ABB RAPID module: Module1.mod

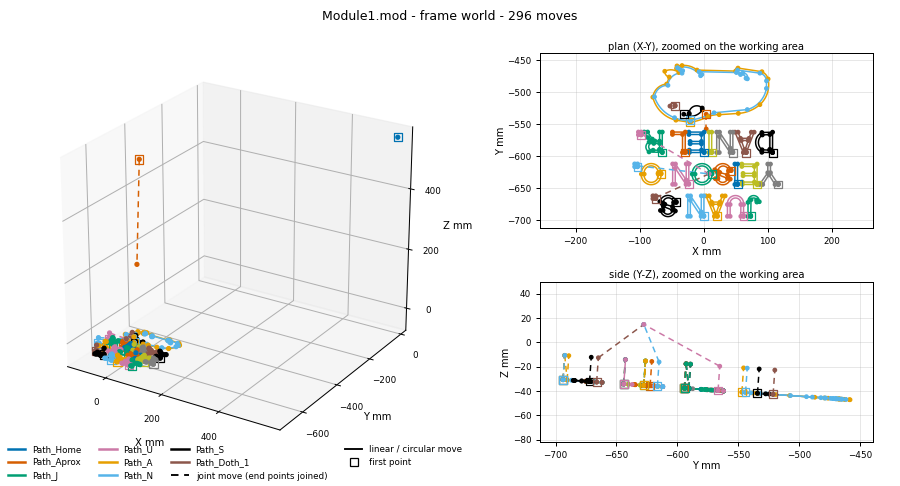
[picture p0: tool path of Module1.mod in frame world, 296 of 313 moves have a stored position in this frame; points joined in program order, loops and branches not executed]
MODULE Module1
    PERS tooldata Tool_Cuy:=[TRUE,[[59.512,0,113],[0.866025404,0,0.5,0]],[1,[0,0,1],[1,0,0,0],0,0,0]];
    TASK PERS wobjdata Workobject_1:=[FALSE,TRUE,"",[[0,-210.462735229,0],[1,0,0,0]],[[-172,-492.000264771,-30],[0.024677671,0.706676031,0.706676031,-0.024677671]]];
    CONST robtarget Target_Aprox:=[[126.462735229,176,-601],[0.999847695,0,0.017452406,0],[0,0,0,0],[9E+09,9E+09,9E+09,9E+09,9E+09,9E+09]];
    CONST robtarget Target_Aprox_2:=[[126.462735229,176,-271],[0.999847695,0,0.017452406,0],[-1,0,-1,1],[9E+09,9E+09,9E+09,9E+09,9E+09,9E+09]];
    CONST robtarget Target_10:=[[8.567735229,245.504,0],[1,0,0,0],[-1,0,-1,1],[9E+09,9E+09,9E+09,9E+09,9E+09,9E+09]];
    CONST robtarget Target_20:=[[34.618735229,245.975,0],[1,0,0,0],[-1,0,-1,1],[9E+09,9E+09,9E+09,9E+09,9E+09,9E+09]];
    CONST robtarget Target_30:=[[37.330735229,250.322,0],[1,0,0,0],[-1,0,-1,1],[9E+09,9E+09,9E+09,9E+09,9E+09,9E+09]];
    CONST robtarget Target_40:=[[34.039735229,254.656,0],[1,0,0,0],[-1,0,-1,1],[9E+09,9E+09,9E+09,9E+09,9E+09,9E+09]];
    CONST robtarget Target_50:=[[30.950735229,255.072,0],[1,0,0,0],[-1,0,-1,1],[9E+09,9E+09,9E+09,9E+09,9E+09,9E+09]];
    CONST robtarget Target_60:=[[31.469735229,258.893,0],[1,0,0,0],[-1,0,-1,1],[9E+09,9E+09,9E+09,9E+09,9E+09,9E+09]];
    CONST robtarget Target_70:=[[41.106735229,250.305,0],[1,0,0,0],[-1,0,-1,1],[9E+09,9E+09,9E+09,9E+09,9E+09,9E+09]];
    CONST robtarget Target_80:=[[30.379735229,241.298,0],[1,0,0,0],[-1,0,-1,1],[9E+09,9E+09,9E+09,9E+09,9E+09,9E+09]];
    CONST robtarget Target_90:=[[8.572735229,241.269,0],[1,0,0,0],[-1,0,-1,1],[9E+09,9E+09,9E+09,9E+09,9E+09,9E+09]];
    CONST robtarget Target_100:=[[8.567735229,245.504,-20],[1,0,0,0],[-1,0,-1,1],[9E+09,9E+09,9E+09,9E+09,9E+09,9E+09]];
    CONST robtarget Target_120:=[[27.070735229,234.308,0],[1,0,0,0],[-1,0,-1,1],[9E+09,9E+09,9E+09,9E+09,9E+09,9E+09]];
    CONST robtarget Target_110:=[[8.582735229,234.284,0],[1,0,0,0],[-1,0,-1,1],[9E+09,9E+09,9E+09,9E+09,9E+09,9E+09]];
    CONST robtarget Target_130:=[[41.144735229,221.667,0],[1,0,0,0],[-1,0,-1,1],[9E+09,9E+09,9E+09,9E+09,9E+09,9E+09]];
    CONST robtarget Target_140:=[[27.103735229,209.141,0],[1,0,0,0],[-1,0,-1,1],[9E+09,9E+09,9E+09,9E+09,9E+09,9E+09]];
    CONST robtarget Target_150:=[[8.615735229,209.116,0],[1,0,0,0],[-1,0,-1,1],[9E+09,9E+09,9E+09,9E+09,9E+09,9E+09]];
    CONST robtarget Target_160:=[[8.609735229,213.351,0],[1,0,0,0],[-1,0,-1,1],[9E+09,9E+09,9E+09,9E+09,9E+09,9E+09]];
    CONST robtarget Target_170:=[[27.076735229,213.375,0],[1,0,0,0],[-1,0,-1,1],[9E+09,9E+09,9E+09,9E+09,9E+09,9E+09]];
    CONST robtarget Target_180:=[[37.324735229,222.033,0],[1,0,0,0],[-1,0,-1,1],[9E+09,9E+09,9E+09,9E+09,9E+09,9E+09]];
    CONST robtarget Target_190:=[[27.054735229,230.074,0],[1,0,0,0],[-1,0,-1,1],[9E+09,9E+09,9E+09,9E+09,9E+09,9E+09]];
    CONST robtarget Target_200:=[[8.587735229,230.049,0],[1,0,0,0],[-1,0,-1,1],[9E+09,9E+09,9E+09,9E+09,9E+09,9E+09]];
    CONST robtarget Target_210:=[[8.582735229,234.284,-20],[1,0,0,0],[-1,0,-1,1],[9E+09,9E+09,9E+09,9E+09,9E+09,9E+09]];
    CONST robtarget Target_220:=[[8.636735229,193.291,0],[1,0,0,0],[-1,0,-1,1],[9E+09,9E+09,9E+09,9E+09,9E+09,9E+09]];
    CONST robtarget Target_230:=[[40.619735229,205.622,0],[1,0,0,0],[-1,0,-1,1],[9E+09,9E+09,9E+09,9E+09,9E+09,9E+09]];
    CONST robtarget Target_240:=[[40.625735229,201.126,0],[1,0,0,0],[-1,0,-1,1],[9E+09,9E+09,9E+09,9E+09,9E+09,9E+09]];
    CONST robtarget Target_250:=[[30.938735229,197.599,0],[1,0,0,0],[-1,0,-1,1],[9E+09,9E+09,9E+09,9E+09,9E+09,9E+09]];
    CONST robtarget Target_260:=[[30.956735229,184.218,0],[1,0,0,0],[-1,0,-1,1],[9E+09,9E+09,9E+09,9E+09,9E+09,9E+09]];
    CONST robtarget Target_270:=[[40.653735229,180.498,0],[1,0,0,0],[-1,0,-1,1],[9E+09,9E+09,9E+09,9E+09,9E+09,9E+09]];
    CONST robtarget Target_280:=[[40.659735229,175.674,0],[1,0,0,0],[-1,0,-1,1],[9E+09,9E+09,9E+09,9E+09,9E+09,9E+09]];
    CONST robtarget Target_290:=[[8.642735229,188.729,0],[1,0,0,0],[-1,0,-1,1],[9E+09,9E+09,9E+09,9E+09,9E+09,9E+09]];
    CONST robtarget Target_300:=[[8.636735229,193.291,-20],[1,0,0,0],[-1,0,-1,1],[9E+09,9E+09,9E+09,9E+09,9E+09,9E+09]];
    CONST robtarget Target_310:=[[12.000735229,191.113,0],[1,0,0,0],[-1,0,-1,1],[9E+09,9E+09,9E+09,9E+09,9E+09,9E+09]];
    CONST robtarget Target_320:=[[27.491735229,196.372,0],[1,0,0,0],[-1,0,-1,1],[9E+09,9E+09,9E+09,9E+09,9E+09,9E+09]];
    CONST robtarget Target_330:=[[27.505735229,185.523,0],[1,0,0,0],[-1,0,-1,1],[9E+09,9E+09,9E+09,9E+09,9E+09,9E+09]];
    CONST robtarget Target_340:=[[12.000735229,191.113,-20],[1,0,0,0],[-1,0,-1,1],[9E+09,9E+09,9E+09,9E+09,9E+09,9E+09]];
    CONST robtarget Target_350:=[[8.663735229,172.292,0],[1,0,0,0],[-1,0,-1,1],[9E+09,9E+09,9E+09,9E+09,9E+09,9E+09]];
    CONST robtarget Target_360:=[[40.663735229,172.334,0],[1,0,0,0],[-1,0,-1,1],[9E+09,9E+09,9E+09,9E+09,9E+09,9E+09]];
    CONST robtarget Target_370:=[[40.669735229,168.274,0],[1,0,0,0],[-1,0,-1,1],[9E+09,9E+09,9E+09,9E+09,9E+09,9E+09]];
    CONST robtarget Target_380:=[[15.523735229,168.241,0],[1,0,0,0],[-1,0,-1,1],[9E+09,9E+09,9E+09,9E+09,9E+09,9E+09]];
    CONST robtarget Target_390:=[[40.691735229,151.467,0],[1,0,0,0],[-1,0,-1,1],[9E+09,9E+09,9E+09,9E+09,9E+09,9E+09]];
    CONST robtarget Target_400:=[[40.696735229,147.123,0],[1,0,0,0],[-1,0,-1,1],[9E+09,9E+09,9E+09,9E+09,9E+09,9E+09]];
    CONST robtarget Target_410:=[[8.696735229,147.081,0],[1,0,0,0],[-1,0,-1,1],[9E+09,9E+09,9E+09,9E+09,9E+09,9E+09]];
    CONST robtarget Target_420:=[[8.691735229,151.141,0],[1,0,0,0],[-1,0,-1,1],[9E+09,9E+09,9E+09,9E+09,9E+09,9E+09]];
    CONST robtarget Target_430:=[[33.815735229,151.174,0],[1,0,0,0],[-1,0,-1,1],[9E+09,9E+09,9E+09,9E+09,9E+09,9E+09]];
    CONST robtarget Target_440:=[[8.669735229,167.949,0],[1,0,0,0],[-1,0,-1,1],[9E+09,9E+09,9E+09,9E+09,9E+09,9E+09]];
    CONST robtarget Target_450:=[[8.663735229,172.292,-20],[1,0,0,0],[-1,0,-1,1],[9E+09,9E+09,9E+09,9E+09,9E+09,9E+09]];
    CONST robtarget Target_460:=[[30.439735229,129.014,0],[1,0,0,0],[-1,0,-1,1],[9E+09,9E+09,9E+09,9E+09,9E+09,9E+09]];
    CONST robtarget Target_470:=[[41.284735229,115.386,0],[1,0,0,0],[-1,0,-1,1],[9E+09,9E+09,9E+09,9E+09,9E+09,9E+09]];
    CONST robtarget Target_480:=[[31.717735229,103.542,0],[1,0,0,0],[-1,0,-1,1],[9E+09,9E+09,9E+09,9E+09,9E+09,9E+09]];
    CONST robtarget Target_490:=[[27.164735229,104.868,0],[1,0,0,0],[-1,0,-1,1],[9E+09,9E+09,9E+09,9E+09,9E+09,9E+09]];
    CONST robtarget Target_500:=[[23.895735229,108.989,0],[1,0,0,0],[-1,0,-1,1],[9E+09,9E+09,9E+09,9E+09,9E+09,9E+09]];
    CONST robtarget Target_510:=[[18.288735229,123.383,0],[1,0,0,0],[-1,0,-1,1],[9E+09,9E+09,9E+09,9E+09,9E+09,9E+09]];
    CONST robtarget Target_520:=[[11.924735229,116.329,0],[1,0,0,0],[-1,0,-1,1],[9E+09,9E+09,9E+09,9E+09,9E+09,9E+09]];
    CONST robtarget Target_530:=[[18.068735229,108.545,0],[1,0,0,0],[-1,0,-1,1],[9E+09,9E+09,9E+09,9E+09,9E+09,9E+09]];
    CONST robtarget Target_540:=[[17.768735229,104.484,0],[1,0,0,0],[-1,0,-1,1],[9E+09,9E+09,9E+09,9E+09,9E+09,9E+09]];
    CONST robtarget Target_550:=[[8.191735229,116.499,0],[1,0,0,0],[-1,0,-1,1],[9E+09,9E+09,9E+09,9E+09,9E+09,9E+09]];
    CONST robtarget Target_560:=[[16.995735229,127.774,0],[1,0,0,0],[-1,0,-1,1],[9E+09,9E+09,9E+09,9E+09,9E+09,9E+09]];
    CONST robtarget Target_570:=[[20.980735229,126.655,0],[1,0,0,0],[-1,0,-1,1],[9E+09,9E+09,9E+09,9E+09,9E+09,9E+09]];
    CONST robtarget Target_580:=[[23.964735229,123.243,0],[1,0,0,0],[-1,0,-1,1],[9E+09,9E+09,9E+09,9E+09,9E+09,9E+09]];
    CONST robtarget Target_590:=[[27.538735229,111.373,0],[1,0,0,0],[-1,0,-1,1],[9E+09,9E+09,9E+09,9E+09,9E+09,9E+09]];
    CONST robtarget Target_600:=[[29.429735229,108.494,0],[1,0,0,0],[-1,0,-1,1],[9E+09,9E+09,9E+09,9E+09,9E+09,9E+09]];
    CONST robtarget Target_610:=[[37.486735229,115.577,0],[1,0,0,0],[-1,0,-1,1],[9E+09,9E+09,9E+09,9E+09,9E+09,9E+09]];
    CONST robtarget Target_620:=[[30.095735229,125.019,0],[1,0,0,0],[-1,0,-1,1],[9E+09,9E+09,9E+09,9E+09,9E+09,9E+09]];
    CONST robtarget Target_630:=[[30.439735229,129.014,-20],[1,0,0,0],[-1,0,-1,1],[9E+09,9E+09,9E+09,9E+09,9E+09,9E+09]];
    CONST robtarget Target_680:=[[36.287735229,97.153,-20],[1,0,0,0],[-1,0,-1,1],[9E+09,9E+09,9E+09,9E+09,9E+09,9E+09]];
    CONST robtarget Target_670:=[[36.293735229,92.678,0],[1,0,0,0],[-1,0,-1,1],[9E+09,9E+09,9E+09,9E+09,9E+09,9E+09]];
    CONST robtarget Target_660:=[[40.768735229,92.684,0],[1,0,0,0],[-1,0,-1,1],[9E+09,9E+09,9E+09,9E+09,9E+09,9E+09]];
    CONST robtarget Target_650:=[[40.762735229,97.159,0],[1,0,0,0],[-1,0,-1,1],[9E+09,9E+09,9E+09,9E+09,9E+09,9E+09]];
    CONST robtarget Target_640:=[[36.287735229,97.153,0],[1,0,0,0],[-1,0,-1,1],[9E+09,9E+09,9E+09,9E+09,9E+09,9E+09]];
    CONST robtarget Target_690:=[[58.453735229,288.658,0],[1,0,0,0],[-1,0,-1,1],[9E+09,9E+09,9E+09,9E+09,9E+09,9E+09]];
    CONST robtarget Target_700:=[[76.914735229,276.35,0],[1,0,0,0],[-1,0,-1,1],[9E+09,9E+09,9E+09,9E+09,9E+09,9E+09]];
    CONST robtarget Target_710:=[[90.469735229,276.367,0],[1,0,0,0],[-1,0,-1,1],[9E+09,9E+09,9E+09,9E+09,9E+09,9E+09]];
    CONST robtarget Target_720:=[[90.475735229,272.133,0],[1,0,0,0],[-1,0,-1,1],[9E+09,9E+09,9E+09,9E+09,9E+09,9E+09]];
    CONST robtarget Target_730:=[[76.919735229,272.115,0],[1,0,0,0],[-1,0,-1,1],[9E+09,9E+09,9E+09,9E+09,9E+09,9E+09]];
    CONST robtarget Target_740:=[[58.491735229,259.321,0],[1,0,0,0],[-1,0,-1,1],[9E+09,9E+09,9E+09,9E+09,9E+09,9E+09]];
    CONST robtarget Target_750:=[[58.485735229,264.254,0],[1,0,0,0],[-1,0,-1,1],[9E+09,9E+09,9E+09,9E+09,9E+09,9E+09]];
    CONST robtarget Target_760:=[[73.534735229,273.966,0],[1,0,0,0],[-1,0,-1,1],[9E+09,9E+09,9E+09,9E+09,9E+09,9E+09]];
    CONST robtarget Target_770:=[[58.460735229,283.507,0],[1,0,0,0],[-1,0,-1,1],[9E+09,9E+09,9E+09,9E+09,9E+09,9E+09]];
    CONST robtarget Target_780:=[[58.453735229,288.658,-20],[1,0,0,0],[-1,0,-1,1],[9E+09,9E+09,9E+09,9E+09,9E+09,9E+09]];
    CONST robtarget Target_790:=[[58.497735229,255.436,0],[1,0,0,0],[-1,0,-1,1],[9E+09,9E+09,9E+09,9E+09,9E+09,9E+09]];
    CONST robtarget Target_800:=[[90.497735229,255.478,0],[1,0,0,0],[-1,0,-1,1],[9E+09,9E+09,9E+09,9E+09,9E+09,9E+09]];
    CONST robtarget Target_810:=[[90.528735229,231.598,0],[1,0,0,0],[-1,0,-1,1],[9E+09,9E+09,9E+09,9E+09,9E+09,9E+09]];
    CONST robtarget Target_820:=[[86.752735229,231.593,0],[1,0,0,0],[-1,0,-1,1],[9E+09,9E+09,9E+09,9E+09,9E+09,9E+09]];
    CONST robtarget Target_830:=[[86.726735229,251.238,0],[1,0,0,0],[-1,0,-1,1],[9E+09,9E+09,9E+09,9E+09,9E+09,9E+09]];
    CONST robtarget Target_840:=[[75.834735229,251.224,0],[1,0,0,0],[-1,0,-1,1],[9E+09,9E+09,9E+09,9E+09,9E+09,9E+09]];
    CONST robtarget Target_850:=[[75.857735229,233.521,0],[1,0,0,0],[-1,0,-1,1],[9E+09,9E+09,9E+09,9E+09,9E+09,9E+09]];
    CONST robtarget Target_860:=[[72.103735229,233.516,0],[1,0,0,0],[-1,0,-1,1],[9E+09,9E+09,9E+09,9E+09,9E+09,9E+09]];
    CONST robtarget Target_870:=[[72.079735229,251.219,0],[1,0,0,0],[-1,0,-1,1],[9E+09,9E+09,9E+09,9E+09,9E+09,9E+09]];
    CONST robtarget Target_880:=[[62.278735229,251.206,0],[1,0,0,0],[-1,0,-1,1],[9E+09,9E+09,9E+09,9E+09,9E+09,9E+09]];
    CONST robtarget Target_890:=[[62.303735229,232.303,0],[1,0,0,0],[-1,0,-1,1],[9E+09,9E+09,9E+09,9E+09,9E+09,9E+09]];
    CONST robtarget Target_900:=[[58.527735229,232.298,0],[1,0,0,0],[-1,0,-1,1],[9E+09,9E+09,9E+09,9E+09,9E+09,9E+09]];
    CONST robtarget Target_910:=[[58.497735229,255.436,-20],[1,0,0,0],[-1,0,-1,1],[9E+09,9E+09,9E+09,9E+09,9E+09,9E+09]];
    CONST robtarget Target_920:=[[58.537735229,224.986,0],[1,0,0,0],[-1,0,-1,1],[9E+09,9E+09,9E+09,9E+09,9E+09,9E+09]];
    CONST robtarget Target_930:=[[90.537735229,225.028,0],[1,0,0,0],[-1,0,-1,1],[9E+09,9E+09,9E+09,9E+09,9E+09,9E+09]];
    CONST robtarget Target_940:=[[90.542735229,220.793,0],[1,0,0,0],[-1,0,-1,1],[9E+09,9E+09,9E+09,9E+09,9E+09,9E+09]];
    CONST robtarget Target_950:=[[58.542735229,220.751,0],[1,0,0,0],[-1,0,-1,1],[9E+09,9E+09,9E+09,9E+09,9E+09,9E+09]];
    CONST robtarget Target_960:=[[58.537735229,224.986,-20],[1,0,0,0],[-1,0,-1,1],[9E+09,9E+09,9E+09,9E+09,9E+09,9E+09]];
    CONST robtarget Target_460_2:=[[80.269735229,214.755,0],[1,0,0,0],[-1,0,-1,1],[9E+09,9E+09,9E+09,9E+09,9E+09,9E+09]];
    CONST robtarget Target_470_2:=[[91.114735229,201.127,0],[1,0,0,0],[-1,0,-1,1],[9E+09,9E+09,9E+09,9E+09,9E+09,9E+09]];
    CONST robtarget Target_480_2:=[[81.547735229,189.283,0],[1,0,0,0],[-1,0,-1,1],[9E+09,9E+09,9E+09,9E+09,9E+09,9E+09]];
    CONST robtarget Target_490_2:=[[76.994735229,190.609,0],[1,0,0,0],[-1,0,-1,1],[9E+09,9E+09,9E+09,9E+09,9E+09,9E+09]];
    CONST robtarget Target_500_2:=[[73.725735229,194.73,0],[1,0,0,0],[-1,0,-1,1],[9E+09,9E+09,9E+09,9E+09,9E+09,9E+09]];
    CONST robtarget Target_510_2:=[[68.118735229,209.124,0],[1,0,0,0],[-1,0,-1,1],[9E+09,9E+09,9E+09,9E+09,9E+09,9E+09]];
    CONST robtarget Target_520_2:=[[61.754735229,202.07,0],[1,0,0,0],[-1,0,-1,1],[9E+09,9E+09,9E+09,9E+09,9E+09,9E+09]];
    CONST robtarget Target_530_2:=[[67.898735229,194.286,0],[1,0,0,0],[-1,0,-1,1],[9E+09,9E+09,9E+09,9E+09,9E+09,9E+09]];
    CONST robtarget Target_540_2:=[[67.598735229,190.225,0],[1,0,0,0],[-1,0,-1,1],[9E+09,9E+09,9E+09,9E+09,9E+09,9E+09]];
    CONST robtarget Target_550_2:=[[58.021735229,202.24,0],[1,0,0,0],[-1,0,-1,1],[9E+09,9E+09,9E+09,9E+09,9E+09,9E+09]];
    CONST robtarget Target_560_2:=[[66.825735229,213.515,0],[1,0,0,0],[-1,0,-1,1],[9E+09,9E+09,9E+09,9E+09,9E+09,9E+09]];
    CONST robtarget Target_570_2:=[[70.810735229,212.396,0],[1,0,0,0],[-1,0,-1,1],[9E+09,9E+09,9E+09,9E+09,9E+09,9E+09]];
    CONST robtarget Target_580_2:=[[73.794735229,208.984,0],[1,0,0,0],[-1,0,-1,1],[9E+09,9E+09,9E+09,9E+09,9E+09,9E+09]];
    CONST robtarget Target_590_2:=[[77.368735229,197.114,0],[1,0,0,0],[-1,0,-1,1],[9E+09,9E+09,9E+09,9E+09,9E+09,9E+09]];
    CONST robtarget Target_600_2:=[[79.259735229,194.235,0],[1,0,0,0],[-1,0,-1,1],[9E+09,9E+09,9E+09,9E+09,9E+09,9E+09]];
    CONST robtarget Target_610_2:=[[87.316735229,201.318,0],[1,0,0,0],[-1,0,-1,1],[9E+09,9E+09,9E+09,9E+09,9E+09,9E+09]];
    CONST robtarget Target_620_2:=[[79.925735229,210.76,0],[1,0,0,0],[-1,0,-1,1],[9E+09,9E+09,9E+09,9E+09,9E+09,9E+09]];
    CONST robtarget Target_630_2:=[[80.269735229,214.755,-20],[1,0,0,0],[-1,0,-1,1],[9E+09,9E+09,9E+09,9E+09,9E+09,9E+09]];
    CONST robtarget Target_970:=[[75.004735229,184.778,0],[1,0,0,0],[-1,0,-1,1],[9E+09,9E+09,9E+09,9E+09,9E+09,9E+09]];
    CONST robtarget Target_980:=[[91.155735229,169.498,0],[1,0,0,0],[-1,0,-1,1],[9E+09,9E+09,9E+09,9E+09,9E+09,9E+09]];
    CONST robtarget Target_990:=[[74.674735229,154.175,0],[1,0,0,0],[-1,0,-1,1],[9E+09,9E+09,9E+09,9E+09,9E+09,9E+09]];
    CONST robtarget Target_1000:=[[58.042735229,169.432,0],[1,0,0,0],[-1,0,-1,1],[9E+09,9E+09,9E+09,9E+09,9E+09,9E+09]];
    CONST robtarget Target_1010:=[[75.004735229,184.778,-20],[1,0,0,0],[-1,0,-1,1],[9E+09,9E+09,9E+09,9E+09,9E+09,9E+09]];
    CONST robtarget Target_1020:=[[75.076735229,180.412,0],[1,0,0,0],[-1,0,-1,1],[9E+09,9E+09,9E+09,9E+09,9E+09,9E+09]];
    CONST robtarget Target_1030:=[[87.532735229,169.515,0],[1,0,0,0],[-1,0,-1,1],[9E+09,9E+09,9E+09,9E+09,9E+09,9E+09]];
    CONST robtarget Target_1040:=[[74.646735229,158.54,0],[1,0,0,0],[-1,0,-1,1],[9E+09,9E+09,9E+09,9E+09,9E+09,9E+09]];
    CONST robtarget Target_1050:=[[61.688735229,169.415,0],[1,0,0,0],[-1,0,-1,1],[9E+09,9E+09,9E+09,9E+09,9E+09,9E+09]];
    CONST robtarget Target_1060:=[[75.076735229,180.412,-20],[1,0,0,0],[-1,0,-1,1],[9E+09,9E+09,9E+09,9E+09,9E+09,9E+09]];
    CONST robtarget Target_350_2:=[[58.637735229,148.74,0],[1,0,0,0],[-1,0,-1,1],[9E+09,9E+09,9E+09,9E+09,9E+09,9E+09]];
    CONST robtarget Target_360_2:=[[90.637735229,148.782,0],[1,0,0,0],[-1,0,-1,1],[9E+09,9E+09,9E+09,9E+09,9E+09,9E+09]];
    CONST robtarget Target_370_2:=[[90.643735229,144.722,0],[1,0,0,0],[-1,0,-1,1],[9E+09,9E+09,9E+09,9E+09,9E+09,9E+09]];
    CONST robtarget Target_380_2:=[[65.497735229,144.689,0],[1,0,0,0],[-1,0,-1,1],[9E+09,9E+09,9E+09,9E+09,9E+09,9E+09]];
    CONST robtarget Target_390_2:=[[90.665735229,127.915,0],[1,0,0,0],[-1,0,-1,1],[9E+09,9E+09,9E+09,9E+09,9E+09,9E+09]];
    CONST robtarget Target_400_2:=[[90.670735229,123.571,0],[1,0,0,0],[-1,0,-1,1],[9E+09,9E+09,9E+09,9E+09,9E+09,9E+09]];
    CONST robtarget Target_410_2:=[[58.670735229,123.529,0],[1,0,0,0],[-1,0,-1,1],[9E+09,9E+09,9E+09,9E+09,9E+09,9E+09]];
    CONST robtarget Target_420_2:=[[58.665735229,127.589,0],[1,0,0,0],[-1,0,-1,1],[9E+09,9E+09,9E+09,9E+09,9E+09,9E+09]];
    CONST robtarget Target_430_2:=[[83.789735229,127.622,0],[1,0,0,0],[-1,0,-1,1],[9E+09,9E+09,9E+09,9E+09,9E+09,9E+09]];
    CONST robtarget Target_440_2:=[[58.643735229,144.397,0],[1,0,0,0],[-1,0,-1,1],[9E+09,9E+09,9E+09,9E+09,9E+09,9E+09]];
    CONST robtarget Target_450_2:=[[58.637735229,148.74,-20],[1,0,0,0],[-1,0,-1,1],[9E+09,9E+09,9E+09,9E+09,9E+09,9E+09]];
    CONST robtarget Target_640_2:=[[86.268735229,68.645,0],[1,0,0,0],[-1,0,-1,1],[9E+09,9E+09,9E+09,9E+09,9E+09,9E+09]];
    CONST robtarget Target_650_2:=[[90.743735229,68.651,0],[1,0,0,0],[-1,0,-1,1],[9E+09,9E+09,9E+09,9E+09,9E+09,9E+09]];
    CONST robtarget Target_660_2:=[[90.749735229,64.176,0],[1,0,0,0],[-1,0,-1,1],[9E+09,9E+09,9E+09,9E+09,9E+09,9E+09]];
    CONST robtarget Target_670_2:=[[86.274735229,64.17,0],[1,0,0,0],[-1,0,-1,1],[9E+09,9E+09,9E+09,9E+09,9E+09,9E+09]];
    CONST robtarget Target_680_2:=[[86.268735229,68.645,-20],[1,0,0,0],[-1,0,-1,1],[9E+09,9E+09,9E+09,9E+09,9E+09,9E+09]];
    CONST robtarget Target_970_2:=[[75.109735229,105.302,0],[1,0,0,0],[-1,0,-1,1],[9E+09,9E+09,9E+09,9E+09,9E+09,9E+09]];
    CONST robtarget Target_980_2:=[[91.260735229,90.022,0],[1,0,0,0],[-1,0,-1,1],[9E+09,9E+09,9E+09,9E+09,9E+09,9E+09]];
    CONST robtarget Target_990_2:=[[74.779735229,74.699,0],[1,0,0,0],[-1,0,-1,1],[9E+09,9E+09,9E+09,9E+09,9E+09,9E+09]];
    CONST robtarget Target_1000_2:=[[58.147735229,89.956,0],[1,0,0,0],[-1,0,-1,1],[9E+09,9E+09,9E+09,9E+09,9E+09,9E+09]];
    CONST robtarget Target_1010_2:=[[75.109735229,105.302,-20],[1,0,0,0],[-1,0,-1,1],[9E+09,9E+09,9E+09,9E+09,9E+09,9E+09]];
    CONST robtarget Target_1020_2:=[[75.181735229,100.936,0],[1,0,0,0],[-1,0,-1,1],[9E+09,9E+09,9E+09,9E+09,9E+09,9E+09]];
    CONST robtarget Target_1030_2:=[[87.637735229,90.039,0],[1,0,0,0],[-1,0,-1,1],[9E+09,9E+09,9E+09,9E+09,9E+09,9E+09]];
    CONST robtarget Target_1040_2:=[[74.751735229,79.064,0],[1,0,0,0],[-1,0,-1,1],[9E+09,9E+09,9E+09,9E+09,9E+09,9E+09]];
    CONST robtarget Target_1050_2:=[[61.793735229,89.939,0],[1,0,0,0],[-1,0,-1,1],[9E+09,9E+09,9E+09,9E+09,9E+09,9E+09]];
    CONST robtarget Target_1060_2:=[[75.181735229,100.936,-20],[1,0,0,0],[-1,0,-1,1],[9E+09,9E+09,9E+09,9E+09,9E+09,9E+09]];
    CONST robtarget Target_1070:=[[108.407735229,279.611,0],[1,0,0,0],[-1,0,-1,1],[9E+09,9E+09,9E+09,9E+09,9E+09,9E+09]];
    CONST robtarget Target_1080:=[[140.407735229,279.653,0],[1,0,0,0],[-1,0,-1,1],[9E+09,9E+09,9E+09,9E+09,9E+09,9E+09]];
    CONST robtarget Target_1090:=[[139.884735229,262.964,0],[1,0,0,0],[-1,0,-1,1],[9E+09,9E+09,9E+09,9E+09,9E+09,9E+09]];
    CONST robtarget Target_1100:=[[124.268735229,253.176,0],[1,0,0,0],[-1,0,-1,1],[9E+09,9E+09,9E+09,9E+09,9E+09,9E+09]];
    CONST robtarget Target_1110:=[[108.888735229,262.891,0],[1,0,0,0],[-1,0,-1,1],[9E+09,9E+09,9E+09,9E+09,9E+09,9E+09]];
    CONST robtarget Target_1120:=[[108.407735229,279.611,-20],[1,0,0,0],[-1,0,-1,1],[9E+09,9E+09,9E+09,9E+09,9E+09,9E+09]];
    CONST robtarget Target_1130:=[[112.189735229,275.381,0],[1,0,0,0],[-1,0,-1,1],[9E+09,9E+09,9E+09,9E+09,9E+09,9E+09]];
    CONST robtarget Target_1140:=[[136.637735229,275.413,0],[1,0,0,0],[-1,0,-1,1],[9E+09,9E+09,9E+09,9E+09,9E+09,9E+09]];
    CONST robtarget Target_1150:=[[136.063735229,263.614,0],[1,0,0,0],[-1,0,-1,1],[9E+09,9E+09,9E+09,9E+09,9E+09,9E+09]];
    CONST robtarget Target_1160:=[[124.196735229,257.541,0],[1,0,0,0],[-1,0,-1,1],[9E+09,9E+09,9E+09,9E+09,9E+09,9E+09]];
    CONST robtarget Target_1170:=[[112.860735229,263.18,0],[1,0,0,0],[-1,0,-1,1],[9E+09,9E+09,9E+09,9E+09,9E+09,9E+09]];
    CONST robtarget Target_1180:=[[112.189735229,275.381,-20],[1,0,0,0],[-1,0,-1,1],[9E+09,9E+09,9E+09,9E+09,9E+09,9E+09]];
    CONST robtarget Target_220_2:=[[108.462735229,238.552,0],[1,0,0,0],[-1,0,-1,1],[9E+09,9E+09,9E+09,9E+09,9E+09,9E+09]];
    CONST robtarget Target_230_2:=[[140.445735229,250.883,0],[1,0,0,0],[-1,0,-1,1],[9E+09,9E+09,9E+09,9E+09,9E+09,9E+09]];
    CONST robtarget Target_240_2:=[[140.451735229,246.387,0],[1,0,0,0],[-1,0,-1,1],[9E+09,9E+09,9E+09,9E+09,9E+09,9E+09]];
    CONST robtarget Target_250_2:=[[130.764735229,242.86,0],[1,0,0,0],[-1,0,-1,1],[9E+09,9E+09,9E+09,9E+09,9E+09,9E+09]];
    CONST robtarget Target_260_2:=[[130.782735229,229.479,0],[1,0,0,0],[-1,0,-1,1],[9E+09,9E+09,9E+09,9E+09,9E+09,9E+09]];
    CONST robtarget Target_270_2:=[[140.479735229,225.759,0],[1,0,0,0],[-1,0,-1,1],[9E+09,9E+09,9E+09,9E+09,9E+09,9E+09]];
    CONST robtarget Target_280_2:=[[140.485735229,220.935,0],[1,0,0,0],[-1,0,-1,1],[9E+09,9E+09,9E+09,9E+09,9E+09,9E+09]];
    CONST robtarget Target_290_2:=[[108.468735229,233.99,0],[1,0,0,0],[-1,0,-1,1],[9E+09,9E+09,9E+09,9E+09,9E+09,9E+09]];
    CONST robtarget Target_300_2:=[[108.462735229,238.552,-20],[1,0,0,0],[-1,0,-1,1],[9E+09,9E+09,9E+09,9E+09,9E+09,9E+09]];
    CONST robtarget Target_310_2:=[[111.826735229,236.374,0],[1,0,0,0],[-1,0,-1,1],[9E+09,9E+09,9E+09,9E+09,9E+09,9E+09]];
    CONST robtarget Target_320_2:=[[127.317735229,241.633,0],[1,0,0,0],[-1,0,-1,1],[9E+09,9E+09,9E+09,9E+09,9E+09,9E+09]];
    CONST robtarget Target_330_2:=[[127.331735229,230.784,0],[1,0,0,0],[-1,0,-1,1],[9E+09,9E+09,9E+09,9E+09,9E+09,9E+09]];
    CONST robtarget Target_340_2:=[[111.826735229,236.374,-20],[1,0,0,0],[-1,0,-1,1],[9E+09,9E+09,9E+09,9E+09,9E+09,9E+09]];
    CONST robtarget Target_350_3:=[[108.489735229,217.553,0],[1,0,0,0],[-1,0,-1,1],[9E+09,9E+09,9E+09,9E+09,9E+09,9E+09]];
    CONST robtarget Target_360_3:=[[140.489735229,217.595,0],[1,0,0,0],[-1,0,-1,1],[9E+09,9E+09,9E+09,9E+09,9E+09,9E+09]];
    CONST robtarget Target_370_3:=[[140.495735229,213.535,0],[1,0,0,0],[-1,0,-1,1],[9E+09,9E+09,9E+09,9E+09,9E+09,9E+09]];
    CONST robtarget Target_380_3:=[[115.349735229,213.502,0],[1,0,0,0],[-1,0,-1,1],[9E+09,9E+09,9E+09,9E+09,9E+09,9E+09]];
    CONST robtarget Target_390_3:=[[140.517735229,196.728,0],[1,0,0,0],[-1,0,-1,1],[9E+09,9E+09,9E+09,9E+09,9E+09,9E+09]];
    CONST robtarget Target_400_3:=[[140.522735229,192.384,0],[1,0,0,0],[-1,0,-1,1],[9E+09,9E+09,9E+09,9E+09,9E+09,9E+09]];
    CONST robtarget Target_410_3:=[[108.522735229,192.342,0],[1,0,0,0],[-1,0,-1,1],[9E+09,9E+09,9E+09,9E+09,9E+09,9E+09]];
    CONST robtarget Target_420_3:=[[108.517735229,196.402,0],[1,0,0,0],[-1,0,-1,1],[9E+09,9E+09,9E+09,9E+09,9E+09,9E+09]];
    CONST robtarget Target_430_3:=[[133.641735229,196.435,0],[1,0,0,0],[-1,0,-1,1],[9E+09,9E+09,9E+09,9E+09,9E+09,9E+09]];
    CONST robtarget Target_440_3:=[[108.495735229,213.21,0],[1,0,0,0],[-1,0,-1,1],[9E+09,9E+09,9E+09,9E+09,9E+09,9E+09]];
    CONST robtarget Target_450_3:=[[108.489735229,217.553,-20],[1,0,0,0],[-1,0,-1,1],[9E+09,9E+09,9E+09,9E+09,9E+09,9E+09]];
    CONST robtarget Target_920_2:=[[108.533735229,184.506,0],[1,0,0,0],[-1,0,-1,1],[9E+09,9E+09,9E+09,9E+09,9E+09,9E+09]];
    CONST robtarget Target_930_2:=[[140.533735229,184.548,0],[1,0,0,0],[-1,0,-1,1],[9E+09,9E+09,9E+09,9E+09,9E+09,9E+09]];
    CONST robtarget Target_940_2:=[[140.538735229,180.313,0],[1,0,0,0],[-1,0,-1,1],[9E+09,9E+09,9E+09,9E+09,9E+09,9E+09]];
    CONST robtarget Target_950_2:=[[108.538735229,180.271,0],[1,0,0,0],[-1,0,-1,1],[9E+09,9E+09,9E+09,9E+09,9E+09,9E+09]];
    CONST robtarget Target_960_2:=[[108.533735229,184.506,-20],[1,0,0,0],[-1,0,-1,1],[9E+09,9E+09,9E+09,9E+09,9E+09,9E+09]];
    CONST robtarget Target_790_2:=[[108.548735229,172.718,0],[1,0,0,0],[-1,0,-1,1],[9E+09,9E+09,9E+09,9E+09,9E+09,9E+09]];
    CONST robtarget Target_800_2:=[[140.548735229,172.76,0],[1,0,0,0],[-1,0,-1,1],[9E+09,9E+09,9E+09,9E+09,9E+09,9E+09]];
    CONST robtarget Target_810_2:=[[140.579735229,148.88,0],[1,0,0,0],[-1,0,-1,1],[9E+09,9E+09,9E+09,9E+09,9E+09,9E+09]];
    CONST robtarget Target_820_2:=[[136.803735229,148.875,0],[1,0,0,0],[-1,0,-1,1],[9E+09,9E+09,9E+09,9E+09,9E+09,9E+09]];
    CONST robtarget Target_830_2:=[[136.777735229,168.52,0],[1,0,0,0],[-1,0,-1,1],[9E+09,9E+09,9E+09,9E+09,9E+09,9E+09]];
    CONST robtarget Target_840_2:=[[125.885735229,168.506,0],[1,0,0,0],[-1,0,-1,1],[9E+09,9E+09,9E+09,9E+09,9E+09,9E+09]];
    CONST robtarget Target_850_2:=[[125.908735229,150.803,0],[1,0,0,0],[-1,0,-1,1],[9E+09,9E+09,9E+09,9E+09,9E+09,9E+09]];
    CONST robtarget Target_860_2:=[[122.154735229,150.798,0],[1,0,0,0],[-1,0,-1,1],[9E+09,9E+09,9E+09,9E+09,9E+09,9E+09]];
    CONST robtarget Target_870_2:=[[122.130735229,168.501,0],[1,0,0,0],[-1,0,-1,1],[9E+09,9E+09,9E+09,9E+09,9E+09,9E+09]];
    CONST robtarget Target_880_2:=[[112.329735229,168.488,0],[1,0,0,0],[-1,0,-1,1],[9E+09,9E+09,9E+09,9E+09,9E+09,9E+09]];
    CONST robtarget Target_890_2:=[[112.354735229,149.585,0],[1,0,0,0],[-1,0,-1,1],[9E+09,9E+09,9E+09,9E+09,9E+09,9E+09]];
    CONST robtarget Target_900_2:=[[108.578735229,149.58,0],[1,0,0,0],[-1,0,-1,1],[9E+09,9E+09,9E+09,9E+09,9E+09,9E+09]];
    CONST robtarget Target_910_2:=[[108.548735229,172.718,-20],[1,0,0,0],[-1,0,-1,1],[9E+09,9E+09,9E+09,9E+09,9E+09,9E+09]];
    CONST robtarget Target_1190:=[[108.587735229,143.163,0],[1,0,0,0],[-1,0,-1,1],[9E+09,9E+09,9E+09,9E+09,9E+09,9E+09]];
    CONST robtarget Target_1200:=[[140.587735229,143.205,0],[1,0,0,0],[-1,0,-1,1],[9E+09,9E+09,9E+09,9E+09,9E+09,9E+09]];
    CONST robtarget Target_1210:=[[140.613735229,123.211,0],[1,0,0,0],[-1,0,-1,1],[9E+09,9E+09,9E+09,9E+09,9E+09,9E+09]];
    CONST robtarget Target_1220:=[[136.837735229,123.206,0],[1,0,0,0],[-1,0,-1,1],[9E+09,9E+09,9E+09,9E+09,9E+09,9E+09]];
    CONST robtarget Target_1230:=[[136.816735229,138.966,0],[1,0,0,0],[-1,0,-1,1],[9E+09,9E+09,9E+09,9E+09,9E+09,9E+09]];
    CONST robtarget Target_1240:=[[108.593735229,138.929,0],[1,0,0,0],[-1,0,-1,1],[9E+09,9E+09,9E+09,9E+09,9E+09,9E+09]];
    CONST robtarget Target_1250:=[[108.587735229,143.163,-20],[1,0,0,0],[-1,0,-1,1],[9E+09,9E+09,9E+09,9E+09,9E+09,9E+09]];
    CONST robtarget Target_1260:=[[108.634735229,107.3,0],[1,0,0,0],[-1,0,-1,1],[9E+09,9E+09,9E+09,9E+09,9E+09,9E+09]];
    CONST robtarget Target_1270:=[[140.634735229,107.342,0],[1,0,0,0],[-1,0,-1,1],[9E+09,9E+09,9E+09,9E+09,9E+09,9E+09]];
    CONST robtarget Target_1280:=[[140.640735229,103.107,0],[1,0,0,0],[-1,0,-1,1],[9E+09,9E+09,9E+09,9E+09,9E+09,9E+09]];
    CONST robtarget Target_1290:=[[126.430735229,103.088,0],[1,0,0,0],[-1,0,-1,1],[9E+09,9E+09,9E+09,9E+09,9E+09,9E+09]];
    CONST robtarget Target_1300:=[[126.592735229,95.82,0],[1,0,0,0],[-1,0,-1,1],[9E+09,9E+09,9E+09,9E+09,9E+09,9E+09]];
    CONST robtarget Target_1310:=[[127.446735229,93.889,0],[1,0,0,0],[-1,0,-1,1],[9E+09,9E+09,9E+09,9E+09,9E+09,9E+09]];
    CONST robtarget Target_1320:=[[129.588735229,91.742,0],[1,0,0,0],[-1,0,-1,1],[9E+09,9E+09,9E+09,9E+09,9E+09,9E+09]];
    CONST robtarget Target_1330:=[[140.664735229,84.466,0],[1,0,0,0],[-1,0,-1,1],[9E+09,9E+09,9E+09,9E+09,9E+09,9E+09]];
    CONST robtarget Target_1340:=[[140.671735229,79.14,0],[1,0,0,0],[-1,0,-1,1],[9E+09,9E+09,9E+09,9E+09,9E+09,9E+09]];
    CONST robtarget Target_1350:=[[131.955735229,84.695,0],[1,0,0,0],[-1,0,-1,1],[9E+09,9E+09,9E+09,9E+09,9E+09,9E+09]];
    CONST robtarget Target_1360:=[[127.694735229,88.203,0],[1,0,0,0],[-1,0,-1,1],[9E+09,9E+09,9E+09,9E+09,9E+09,9E+09]];
    CONST robtarget Target_1370:=[[126.097735229,90.755,0],[1,0,0,0],[-1,0,-1,1],[9E+09,9E+09,9E+09,9E+09,9E+09,9E+09]];
    CONST robtarget Target_1380:=[[125.043735229,86.748,0],[1,0,0,0],[-1,0,-1,1],[9E+09,9E+09,9E+09,9E+09,9E+09,9E+09]];
    CONST robtarget Target_1390:=[[117.399735229,81.729,0],[1,0,0,0],[-1,0,-1,1],[9E+09,9E+09,9E+09,9E+09,9E+09,9E+09]];
    CONST robtarget Target_1400:=[[109.524735229,86.608,0],[1,0,0,0],[-1,0,-1,1],[9E+09,9E+09,9E+09,9E+09,9E+09,9E+09]];
    CONST robtarget Target_1410:=[[108.634735229,107.3,-20],[1,0,0,0],[-1,0,-1,1],[9E+09,9E+09,9E+09,9E+09,9E+09,9E+09]];
    CONST robtarget Target_1420:=[[112.176735229,103.07,0],[1,0,0,0],[-1,0,-1,1],[9E+09,9E+09,9E+09,9E+09,9E+09,9E+09]];
    CONST robtarget Target_1430:=[[122.763735229,103.084,0],[1,0,0,0],[-1,0,-1,1],[9E+09,9E+09,9E+09,9E+09,9E+09,9E+09]];
    CONST robtarget Target_1440:=[[122.775735229,93.981,0],[1,0,0,0],[-1,0,-1,1],[9E+09,9E+09,9E+09,9E+09,9E+09,9E+09]];
    CONST robtarget Target_1450:=[[117.394735229,86.094,0],[1,0,0,0],[-1,0,-1,1],[9E+09,9E+09,9E+09,9E+09,9E+09,9E+09]];
    CONST robtarget Target_1460:=[[112.189735229,92.942,0],[1,0,0,0],[-1,0,-1,1],[9E+09,9E+09,9E+09,9E+09,9E+09,9E+09]];
    CONST robtarget Target_1470:=[[112.176735229,103.07,-20],[1,0,0,0],[-1,0,-1,1],[9E+09,9E+09,9E+09,9E+09,9E+09,9E+09]];
    CONST robtarget Target_640_3:=[[136.203735229,74.507,0],[1,0,0,0],[-1,0,-1,1],[9E+09,9E+09,9E+09,9E+09,9E+09,9E+09]];
    CONST robtarget Target_650_3:=[[140.678735229,74.513,0],[1,0,0,0],[-1,0,-1,1],[9E+09,9E+09,9E+09,9E+09,9E+09,9E+09]];
    CONST robtarget Target_660_3:=[[140.684735229,70.038,0],[1,0,0,0],[-1,0,-1,1],[9E+09,9E+09,9E+09,9E+09,9E+09,9E+09]];
    CONST robtarget Target_670_3:=[[136.209735229,70.032,0],[1,0,0,0],[-1,0,-1,1],[9E+09,9E+09,9E+09,9E+09,9E+09,9E+09]];
    CONST robtarget Target_680_3:=[[136.203735229,74.507,-20],[1,0,0,0],[-1,0,-1,1],[9E+09,9E+09,9E+09,9E+09,9E+09,9E+09]];
    CONST robtarget Target_1480:=[[155.805735229,151.181,0],[1,0,0,0],[-1,0,-1,1],[9E+09,9E+09,9E+09,9E+09,9E+09,9E+09]];
    CONST robtarget Target_1490:=[[159.328735229,165.416,0],[1,0,0,0],[-1,0,-1,1],[9E+09,9E+09,9E+09,9E+09,9E+09,9E+09]];
    CONST robtarget Target_1500:=[[164.805735229,179.181,0],[1,0,0,0],[-1,0,-1,1],[9E+09,9E+09,9E+09,9E+09,9E+09,9E+09]];
    CONST robtarget Target_1510:=[[167.565735229,189.992,0],[1,0,0,0],[-1,0,-1,1],[9E+09,9E+09,9E+09,9E+09,9E+09,9E+09]];
    CONST robtarget Target_1520:=[[167.805735229,196.181,0],[1,0,0,0],[-1,0,-1,1],[9E+09,9E+09,9E+09,9E+09,9E+09,9E+09]];
    CONST robtarget Target_1530:=[[169.805735229,226.181,0],[1,0,0,0],[-1,0,-1,1],[9E+09,9E+09,9E+09,9E+09,9E+09,9E+09]];
    CONST robtarget Target_1540:=[[173.194735229,242.201,0],[1,0,0,0],[-1,0,-1,1],[9E+09,9E+09,9E+09,9E+09,9E+09,9E+09]];
    CONST robtarget Target_1550:=[[183.545735229,259.86,0],[1,0,0,0],[-1,0,-1,1],[9E+09,9E+09,9E+09,9E+09,9E+09,9E+09]];
    CONST robtarget Target_1560:=[[203.805735229,272.181,0],[1,0,0,0],[-1,0,-1,1],[9E+09,9E+09,9E+09,9E+09,9E+09,9E+09]];
    CONST robtarget Target_1570:=[[140.423735229,268.106,0],[1,0,0,0],[-1,0,-1,1],[9E+09,9E+09,9E+09,9E+09,9E+09,9E+09]];
    CONST robtarget Target_1580:=[[223.728735229,272.681,0],[1,0,0,0],[-1,0,-1,1],[9E+09,9E+09,9E+09,9E+09,9E+09,9E+09]];
    CONST robtarget Target_1590:=[[230.071735229,269.481,0],[1,0,0,0],[-1,0,-1,1],[9E+09,9E+09,9E+09,9E+09,9E+09,9E+09]];
    CONST robtarget Target_1600:=[[235.153735229,262.985,0],[1,0,0,0],[-1,0,-1,1],[9E+09,9E+09,9E+09,9E+09,9E+09,9E+09]];
    CONST robtarget Target_1610:=[[240.805735229,225.616,0],[1,0,0,0],[-1,0,-1,1],[9E+09,9E+09,9E+09,9E+09,9E+09,9E+09]];
    CONST robtarget Target_1620:=[[239.305735229,221.948,0],[1,0,0,0],[-1,0,-1,1],[9E+09,9E+09,9E+09,9E+09,9E+09,9E+09]];
    CONST robtarget Target_1630:=[[140.485735229,220.935,0],[1,0,0,0],[-1,0,-1,1],[9E+09,9E+09,9E+09,9E+09,9E+09,9E+09]];
    CONST robtarget Target_1640:=[[236.070735229,221.948,0],[1,0,0,0],[-1,0,-1,1],[9E+09,9E+09,9E+09,9E+09,9E+09,9E+09]];
    CONST robtarget Target_1650:=[[237.687735229,161.589,0],[1,0,0,0],[-1,0,-1,1],[9E+09,9E+09,9E+09,9E+09,9E+09,9E+09]];
    CONST robtarget Target_1660:=[[243.925735229,149.655,0],[1,0,0,0],[-1,0,-1,1],[9E+09,9E+09,9E+09,9E+09,9E+09,9E+09]];
    CONST robtarget Target_1670:=[[244.805735229,138.181,0],[1,0,0,0],[-1,0,-1,1],[9E+09,9E+09,9E+09,9E+09,9E+09,9E+09]];
    CONST robtarget Target_1680:=[[244.215735229,130.298,0],[1,0,0,0],[-1,0,-1,1],[9E+09,9E+09,9E+09,9E+09,9E+09,9E+09]];
    CONST robtarget Target_1690:=[[242.835735229,128.191,0],[1,0,0,0],[-1,0,-1,1],[9E+09,9E+09,9E+09,9E+09,9E+09,9E+09]];
    CONST robtarget Target_1700:=[[239.976735229,129.616,0],[1,0,0,0],[-1,0,-1,1],[9E+09,9E+09,9E+09,9E+09,9E+09,9E+09]];
    CONST robtarget Target_1710:=[[235.981735229,134.906,0],[1,0,0,0],[-1,0,-1,1],[9E+09,9E+09,9E+09,9E+09,9E+09,9E+09]];
    CONST robtarget Target_1720:=[[233.805735229,133.181,0],[1,0,0,0],[-1,0,-1,1],[9E+09,9E+09,9E+09,9E+09,9E+09,9E+09]];
    CONST robtarget Target_1730:=[[237.456735229,125.779,0],[1,0,0,0],[-1,0,-1,1],[9E+09,9E+09,9E+09,9E+09,9E+09,9E+09]];
    CONST robtarget Target_1740:=[[235.805735229,111.181,0],[1,0,0,0],[-1,0,-1,1],[9E+09,9E+09,9E+09,9E+09,9E+09,9E+09]];
    CONST robtarget Target_1750:=[[231.009735229,112.354,0],[1,0,0,0],[-1,0,-1,1],[9E+09,9E+09,9E+09,9E+09,9E+09,9E+09]];
    CONST robtarget Target_1760:=[[226.805735229,118.181,0],[1,0,0,0],[-1,0,-1,1],[9E+09,9E+09,9E+09,9E+09,9E+09,9E+09]];
    CONST robtarget Target_1770:=[[215.805735229,114.181,0],[1,0,0,0],[-1,0,-1,1],[9E+09,9E+09,9E+09,9E+09,9E+09,9E+09]];
    CONST robtarget Target_1780:=[[210.368735229,100.781,0],[1,0,0,0],[-1,0,-1,1],[9E+09,9E+09,9E+09,9E+09,9E+09,9E+09]];
    CONST robtarget Target_1790:=[[195.213735229,92.561,0],[1,0,0,0],[-1,0,-1,1],[9E+09,9E+09,9E+09,9E+09,9E+09,9E+09]];
    CONST robtarget Target_1800:=[[179.805735229,99.181,0],[1,0,0,0],[-1,0,-1,1],[9E+09,9E+09,9E+09,9E+09,9E+09,9E+09]];
    CONST robtarget Target_1810:=[[159.213735229,128.627,0],[1,0,0,0],[-1,0,-1,1],[9E+09,9E+09,9E+09,9E+09,9E+09,9E+09]];
    CONST robtarget Target_1820:=[[155.805735229,151.181,-20],[1,0,0,0],[-1,0,-1,1],[9E+09,9E+09,9E+09,9E+09,9E+09,9E+09]];
    CONST robtarget Target_1830:=[[158.805735229,151.181,0],[1,0,0,0],[-1,0,-1,1],[9E+09,9E+09,9E+09,9E+09,9E+09,9E+09]];
    CONST robtarget Target_1840:=[[164.161735229,171.133,0],[1,0,0,0],[-1,0,-1,1],[9E+09,9E+09,9E+09,9E+09,9E+09,9E+09]];
    CONST robtarget Target_1850:=[[170.805735229,188.181,0],[1,0,0,0],[-1,0,-1,1],[9E+09,9E+09,9E+09,9E+09,9E+09,9E+09]];
    CONST robtarget Target_1860:=[[175.805735229,240.181,0],[1,0,0,0],[-1,0,-1,1],[9E+09,9E+09,9E+09,9E+09,9E+09,9E+09]];
    CONST robtarget Target_1870:=[[184.865735229,256.66,0],[1,0,0,0],[-1,0,-1,1],[9E+09,9E+09,9E+09,9E+09,9E+09,9E+09]];
    CONST robtarget Target_1880:=[[208.939735229,270.031,0],[1,0,0,0],[-1,0,-1,1],[9E+09,9E+09,9E+09,9E+09,9E+09,9E+09]];
    CONST robtarget Target_1890:=[[140.423735229,268.106,0],[1,0,0,0],[-1,0,-1,1],[9E+09,9E+09,9E+09,9E+09,9E+09,9E+09]];
    CONST robtarget Target_1900:=[[220.805735229,270.181,0],[1,0,0,0],[-1,0,-1,1],[9E+09,9E+09,9E+09,9E+09,9E+09,9E+09]];
    CONST robtarget Target_1910:=[[228.236735229,267.216,0],[1,0,0,0],[-1,0,-1,1],[9E+09,9E+09,9E+09,9E+09,9E+09,9E+09]];
    CONST robtarget Target_1920:=[[232.858735229,259.897,0],[1,0,0,0],[-1,0,-1,1],[9E+09,9E+09,9E+09,9E+09,9E+09,9E+09]];
    CONST robtarget Target_1930:=[[237.638735229,224.921,0],[1,0,0,0],[-1,0,-1,1],[9E+09,9E+09,9E+09,9E+09,9E+09,9E+09]];
    CONST robtarget Target_1940:=[[234.665735229,226.928,0],[1,0,0,0],[-1,0,-1,1],[9E+09,9E+09,9E+09,9E+09,9E+09,9E+09]];
    CONST robtarget Target_1950:=[[232.989735229,233.237,0],[1,0,0,0],[-1,0,-1,1],[9E+09,9E+09,9E+09,9E+09,9E+09,9E+09]];
    CONST robtarget Target_1960:=[[229.293735229,239.949,0],[1,0,0,0],[-1,0,-1,1],[9E+09,9E+09,9E+09,9E+09,9E+09,9E+09]];
    CONST robtarget Target_1970:=[[223.971735229,240.28,0],[1,0,0,0],[-1,0,-1,1],[9E+09,9E+09,9E+09,9E+09,9E+09,9E+09]];
    CONST robtarget Target_1980:=[[224.805735229,238.181,0],[1,0,0,0],[-1,0,-1,1],[9E+09,9E+09,9E+09,9E+09,9E+09,9E+09]];
    CONST robtarget Target_1990:=[[226.838735229,237.926,0],[1,0,0,0],[-1,0,-1,1],[9E+09,9E+09,9E+09,9E+09,9E+09,9E+09]];
    CONST robtarget Target_2000:=[[229.805735229,234.681,0],[1,0,0,0],[-1,0,-1,1],[9E+09,9E+09,9E+09,9E+09,9E+09,9E+09]];
    CONST robtarget Target_2010:=[[230.709735229,229.564,0],[1,0,0,0],[-1,0,-1,1],[9E+09,9E+09,9E+09,9E+09,9E+09,9E+09]];
    CONST robtarget Target_2020:=[[233.805735229,223.181,0],[1,0,0,0],[-1,0,-1,1],[9E+09,9E+09,9E+09,9E+09,9E+09,9E+09]];
    CONST robtarget Target_2030:=[[140.548735229,172.761,0],[1,0,0,0],[-1,0,-1,1],[9E+09,9E+09,9E+09,9E+09,9E+09,9E+09]];
    CONST robtarget Target_2040:=[[235.176735229,164.914,0],[1,0,0,0],[-1,0,-1,1],[9E+09,9E+09,9E+09,9E+09,9E+09,9E+09]];
    CONST robtarget Target_2050:=[[233.424735229,167.032,0],[1,0,0,0],[-1,0,-1,1],[9E+09,9E+09,9E+09,9E+09,9E+09,9E+09]];
    CONST robtarget Target_2060:=[[230.805735229,169.181,0],[1,0,0,0],[-1,0,-1,1],[9E+09,9E+09,9E+09,9E+09,9E+09,9E+09]];
    CONST robtarget Target_2070:=[[140.548735229,172.761,0],[1,0,0,0],[-1,0,-1,1],[9E+09,9E+09,9E+09,9E+09,9E+09,9E+09]];
    CONST robtarget Target_2080:=[[228.805735229,167.181,0],[1,0,0,0],[-1,0,-1,1],[9E+09,9E+09,9E+09,9E+09,9E+09,9E+09]];
    CONST robtarget Target_2090:=[[241.565735229,147.814,0],[1,0,0,0],[-1,0,-1,1],[9E+09,9E+09,9E+09,9E+09,9E+09,9E+09]];
    CONST robtarget Target_2100:=[[241.427735229,130.997,0],[1,0,0,0],[-1,0,-1,1],[9E+09,9E+09,9E+09,9E+09,9E+09,9E+09]];
    CONST robtarget Target_2110:=[[238.405735229,135.006,0],[1,0,0,0],[-1,0,-1,1],[9E+09,9E+09,9E+09,9E+09,9E+09,9E+09]];
    CONST robtarget Target_2120:=[[236.805735229,139.181,0],[1,0,0,0],[-1,0,-1,1],[9E+09,9E+09,9E+09,9E+09,9E+09,9E+09]];
    CONST robtarget Target_2130:=[[234.052735229,139.426,0],[1,0,0,0],[-1,0,-1,1],[9E+09,9E+09,9E+09,9E+09,9E+09,9E+09]];
    CONST robtarget Target_2140:=[[232.805735229,138.181,0],[1,0,0,0],[-1,0,-1,1],[9E+09,9E+09,9E+09,9E+09,9E+09,9E+09]];
    CONST robtarget Target_2150:=[[227.651735229,122.877,0],[1,0,0,0],[-1,0,-1,1],[9E+09,9E+09,9E+09,9E+09,9E+09,9E+09]];
    CONST robtarget Target_2160:=[[213.805735229,116.181,0],[1,0,0,0],[-1,0,-1,1],[9E+09,9E+09,9E+09,9E+09,9E+09,9E+09]];
    CONST robtarget Target_2170:=[[211.295735229,105.803,0],[1,0,0,0],[-1,0,-1,1],[9E+09,9E+09,9E+09,9E+09,9E+09,9E+09]];
    CONST robtarget Target_2180:=[[195.805735229,95.181,0],[1,0,0,0],[-1,0,-1,1],[9E+09,9E+09,9E+09,9E+09,9E+09,9E+09]];
    CONST robtarget Target_2190:=[[173.805735229,109.181,0],[1,0,0,0],[-1,0,-1,1],[9E+09,9E+09,9E+09,9E+09,9E+09,9E+09]];
    CONST robtarget Target_2200:=[[163.142735229,126.477,0],[1,0,0,0],[-1,0,-1,1],[9E+09,9E+09,9E+09,9E+09,9E+09,9E+09]];
    CONST robtarget Target_2210:=[[158.805735229,151.181,-20],[1,0,0,0],[-1,0,-1,1],[9E+09,9E+09,9E+09,9E+09,9E+09,9E+09]];
    CONST robtarget Target_2220:=[[159.790735229,137.217,0],[1,0,0,0],[-1,0,-1,1],[9E+09,9E+09,9E+09,9E+09,9E+09,9E+09]];
    CONST robtarget Target_2230:=[[168.537735229,140.909,0],[1,0,0,0],[-1,0,-1,1],[9E+09,9E+09,9E+09,9E+09,9E+09,9E+09]];
    CONST robtarget Target_2240:=[[165.824735229,156.248,0],[1,0,0,0],[-1,0,-1,1],[9E+09,9E+09,9E+09,9E+09,9E+09,9E+09]];
    CONST robtarget Target_2250:=[[175.297735229,169.833,0],[1,0,0,0],[-1,0,-1,1],[9E+09,9E+09,9E+09,9E+09,9E+09,9E+09]];
    CONST robtarget Target_2260:=[[176.805735229,170.181,0],[1,0,0,0],[-1,0,-1,1],[9E+09,9E+09,9E+09,9E+09,9E+09,9E+09]];
    CONST robtarget Target_2270:=[[178.203735229,169.693,0],[1,0,0,0],[-1,0,-1,1],[9E+09,9E+09,9E+09,9E+09,9E+09,9E+09]];
    CONST robtarget Target_2280:=[[180.831735229,156.598,0],[1,0,0,0],[-1,0,-1,1],[9E+09,9E+09,9E+09,9E+09,9E+09,9E+09]];
    CONST robtarget Target_2290:=[[168.641735229,149.303,0],[1,0,0,0],[-1,0,-1,1],[9E+09,9E+09,9E+09,9E+09,9E+09,9E+09]];
    CONST robtarget Target_2300:=[[168.641735229,149.303,-20],[1,0,0,0],[-1,0,-1,1],[9E+09,9E+09,9E+09,9E+09,9E+09,9E+09]];
    CONST robtarget Target_2350:=[[181.505735229,127.281,-20],[1,0,0,0],[-1,0,-1,1],[9E+09,9E+09,9E+09,9E+09,9E+09,9E+09]];
    CONST robtarget Target_2340:=[[177.505735229,123.301,0],[1,0,0,0],[-1,0,-1,1],[9E+09,9E+09,9E+09,9E+09,9E+09,9E+09]];
    CONST robtarget Target_2330:=[[181.248735229,119.29,0],[1,0,0,0],[-1,0,-1,1],[9E+09,9E+09,9E+09,9E+09,9E+09,9E+09]];
    CONST robtarget Target_2320:=[[185.505735229,123.235,0],[1,0,0,0],[-1,0,-1,1],[9E+09,9E+09,9E+09,9E+09,9E+09,9E+09]];
    CONST robtarget Target_2310:=[[181.506735229,127.281,0],[1,0,0,0],[-1,0,-1,1],[9E+09,9E+09,9E+09,9E+09,9E+09,9E+09]];
    CONST jointtarget Aura_Vertical := [[0,-20,20,0,70,0],[9E+09,9E+09,9E+09,9E+09,9E+09,9E+09]];

    CONST jointtarget Aura_Abre_Der := [[10,-40,-20,35,80,-45],[9E+09,9E+09,9E+09,9E+09,9E+09,9E+09]];

    CONST jointtarget Aura_Abre_Izq := [[-10,-20,-10,-35,0,45],[9E+09,9E+09,9E+09,9E+09,9E+09,9E+09]];

    CONST jointtarget Aura_Giro_Der := [[2,10,5,-20,70,-80],[9E+09,9E+09,9E+09,9E+09,9E+09,9E+09]];

    CONST jointtarget Aura_Giro_Izq := [[-2,10,5,0,70,80],[9E+09,9E+09,9E+09,9E+09,9E+09,9E+09]];

    CONST jointtarget Aura_Saludo_1 := [[0,-20,30,0,-30,0],[9E+09,9E+09,9E+09,9E+09,9E+09,9E+09]];
    CONST jointtarget Aura_Saludo_2 := [[0,-20,30,0,20,60],[9E+09,9E+09,9E+09,9E+09,9E+09,9E+09]];
    CONST jointtarget Aura_Saludo_3 := [[0,-20,30,0,-30,120],[9E+09,9E+09,9E+09,9E+09,9E+09,9E+09]];
    CONST jointtarget Aura_Saludo_4 := [[0,-20,30,0,20,180],[9E+09,9E+09,9E+09,9E+09,9E+09,9E+09]];
    CONST jointtarget Aura_Saludo_5 := [[0,-20,30,0,-30,240],[9E+09,9E+09,9E+09,9E+09,9E+09,9E+09]];
    CONST jointtarget Aura_Saludo_6 := [[0,-20,30,0,20,300],[9E+09,9E+09,9E+09,9E+09,9E+09,9E+09]];
    CONST jointtarget Aura_Saludo_Fin := [[0,-20,30,0,-30,0],[9E+09,9E+09,9E+09,9E+09,9E+09,9E+09]];
    CONST jointtarget Mant_Aprox := [[0,-6,27,2,-52,165.75],[9E+09,9E+09,9E+09,9E+09,9E+09,9E+09]];
    CONST robtarget Target_Home:=[[574.396521874,0,571.46109617],[0,0,1,0],[0,0,0,0],[9E+09,9E+09,9E+09,9E+09,9E+09,9E+09]];
    CONST robtarget Target_1020_3:=[[71.588911511,180.412,-49.878202511],[1,0,0,0],[-1,0,-1,1],[9E+09,9E+09,9E+09,9E+09,9E+09,9E+09]];

    PROC main()
        SET FWD_Conveyor;

        WHILE TRUE DO

            IF DI_01 = 1 THEN
                SET BWD_Conveyor;
                WaitTime 3;
                RESET BWD_Conveyor;
                WaitTime 0.5;
                SET DO_01;
                EscribirNombres;
                RESET DO_01;
                SET BWD_Conveyor;
                WaitTime 2;
                RESET BWD_Conveyor;

            ELSEIF DI_01 = 1 AND DI_02 = 1 THEN

                RESET FWD_Conveyor;
                SET BWD_Conveyor;
                WaitTime 5.5;
                RESET BWD_Conveyor;

            ELSEIF DI_03 = 1 THEN
                FarmearAura;
                WaitDI DI_03,0;

            ELSEIF DI_02 = 1 THEN
                Mantenimiento;
                WaitDI DI_02,0;

            ELSE
                WaitTime 0.05;
            ENDIF

        ENDWHILE

    ENDPROC

    PROC EscribirNombres()

            Path_Home;
            Path_Aprox;
            Path_J;
            Path_U;
            Path_A;
            Path_N;
            Path_S;
            Path_Doth_1;
            Path_Y;
            Path_E;
            Path_I;
            Path_S_2;
            Path_O;
            Path_N_2;
            Path_O_2;
            Path_Doth_2;
            Path_D;
            Path_A_2;
            Path_N_3;
            Path_I_2;
            Path_E_2;
            Path_L;
            Path_R;
            Path_Doth_3;
            Path_Cuy_Externo;
            Path_Cuy_Interno;
            Path_Oreja;
            Path_Ojo;
            Path_Home;

    ENDPROC
    PROC Path_Home()
        MoveJ Target_Home,v200,z10,Tool_Cuy\WObj:=wobj0;
    ENDPROC
    PROC Path_Aprox()
        MoveJ Target_Aprox,v200,z10,Tool_Cuy\WObj:=Workobject_1;
        MoveJ Target_Aprox_2,v200,z10,Tool_Cuy\WObj:=Workobject_1;
    ENDPROC
    PROC Path_J()
        MoveJ Target_10,v200,z10,Tool_Cuy\WObj:=Workobject_1;
        MoveL Target_20,v200,z10,Tool_Cuy\WObj:=Workobject_1;
        MoveC Target_30,Target_40,v200,z10,Tool_Cuy\WObj:=Workobject_1;
        MoveL Target_50,v200,z10,Tool_Cuy\WObj:=Workobject_1;
        MoveL Target_60,v200,z10,Tool_Cuy\WObj:=Workobject_1;
        MoveC Target_70,Target_80,v200,z10,Tool_Cuy\WObj:=Workobject_1;
        MoveL Target_90,v200,z10,Tool_Cuy\WObj:=Workobject_1;
        MoveL Target_10,v200,z10,Tool_Cuy\WObj:=Workobject_1;
        MoveJ Target_100,v200,z10,Tool_Cuy\WObj:=Workobject_1;
    ENDPROC
    PROC Path_U()
        MoveJ Target_110,v200,z10,Tool_Cuy\WObj:=Workobject_1;
        MoveL Target_120,v200,z10,Tool_Cuy\WObj:=Workobject_1;
        MoveC Target_130,Target_140,v200,z10,Tool_Cuy\WObj:=Workobject_1;
        MoveL Target_150,v200,z10,Tool_Cuy\WObj:=Workobject_1;
        MoveL Target_160,v200,z10,Tool_Cuy\WObj:=Workobject_1;
        MoveL Target_170,v200,z10,Tool_Cuy\WObj:=Workobject_1;
        MoveC Target_180,Target_190,v200,z10,Tool_Cuy\WObj:=Workobject_1;
        MoveL Target_200,v200,z10,Tool_Cuy\WObj:=Workobject_1;
        MoveL Target_110,v200,z10,Tool_Cuy\WObj:=Workobject_1;
        MoveJ Target_210,v1000,z100,Tool_Cuy\WObj:=Workobject_1;

    ENDPROC
    PROC Path_A()
        MoveJ Target_220,v200,z10,Tool_Cuy\WObj:=Workobject_1;
        MoveL Target_230,v200,z10,Tool_Cuy\WObj:=Workobject_1;
        MoveL Target_240,v200,z10,Tool_Cuy\WObj:=Workobject_1;
        MoveL Target_250,v200,z10,Tool_Cuy\WObj:=Workobject_1;
        MoveL Target_260,v200,z10,Tool_Cuy\WObj:=Workobject_1;
        MoveL Target_270,v200,z10,Tool_Cuy\WObj:=Workobject_1;
        MoveL Target_280,v200,z10,Tool_Cuy\WObj:=Workobject_1;
        MoveL Target_290,v200,z10,Tool_Cuy\WObj:=Workobject_1;
        MoveL Target_220,v200,z10,Tool_Cuy\WObj:=Workobject_1;
        MoveJ Target_300,v200,z10,Tool_Cuy\WObj:=Workobject_1;
        MoveJ Target_310,v200,z10,Tool_Cuy\WObj:=Workobject_1;
        MoveL Target_320,v200,z10,Tool_Cuy\WObj:=Workobject_1;
        MoveL Target_330,v200,z10,Tool_Cuy\WObj:=Workobject_1;
        MoveL Target_310,v200,z10,Tool_Cuy\WObj:=Workobject_1;
        MoveJ Target_340,v200,z10,Tool_Cuy\WObj:=Workobject_1;

    ENDPROC
    PROC Path_N()
        MoveJ Target_350,v200,z10,Tool_Cuy\WObj:=Workobject_1;
        MoveL Target_360,v200,z10,Tool_Cuy\WObj:=Workobject_1;
        MoveL Target_370,v200,z10,Tool_Cuy\WObj:=Workobject_1;
        MoveL Target_380,v200,z10,Tool_Cuy\WObj:=Workobject_1;
        MoveL Target_390,v200,z10,Tool_Cuy\WObj:=Workobject_1;
        MoveL Target_400,v200,z10,Tool_Cuy\WObj:=Workobject_1;
        MoveL Target_410,v200,z10,Tool_Cuy\WObj:=Workobject_1;
        MoveL Target_420,v200,z10,Tool_Cuy\WObj:=Workobject_1;
        MoveL Target_430,v200,z10,Tool_Cuy\WObj:=Workobject_1;
        MoveL Target_440,v200,z10,Tool_Cuy\WObj:=Workobject_1;
        MoveL Target_350,v200,z10,Tool_Cuy\WObj:=Workobject_1;
        MoveJ Target_450,v200,z10,Tool_Cuy\WObj:=Workobject_1;
    ENDPROC
    PROC Path_S()
        MoveJ Target_460,v200,z10,Tool_Cuy\WObj:=Workobject_1;
        MoveC Target_470,Target_480,v200,z10,Tool_Cuy\WObj:=Workobject_1;
        MoveC Target_490,Target_500,v200,z10,Tool_Cuy\WObj:=Workobject_1;
        MoveL Target_510,v200,z10,Tool_Cuy\WObj:=Workobject_1;
        MoveC Target_520,Target_530,v200,z10,Tool_Cuy\WObj:=Workobject_1;
        MoveL Target_540,v200,z10,Tool_Cuy\WObj:=Workobject_1;
        MoveC Target_550,Target_560,v200,z10,Tool_Cuy\WObj:=Workobject_1;
        MoveC Target_570,Target_580,v200,z10,Tool_Cuy\WObj:=Workobject_1;
        MoveL Target_590,v200,z10,Tool_Cuy\WObj:=Workobject_1;
        MoveL Target_600,v200,z10,Tool_Cuy\WObj:=Workobject_1;
        MoveC Target_610,Target_620,v200,z10,Tool_Cuy\WObj:=Workobject_1;
        MoveL Target_460,v200,z10,Tool_Cuy\WObj:=Workobject_1;
        MoveJ Target_630,v200,z10,Tool_Cuy\WObj:=Workobject_1;
    ENDPROC
    PROC Path_Doth_1()
        MoveJ Target_640,v200,z10,Tool_Cuy\WObj:=Workobject_1;
        MoveL Target_650,v200,z10,Tool_Cuy\WObj:=Workobject_1;
        MoveL Target_660,v200,z10,Tool_Cuy\WObj:=Workobject_1;
        MoveL Target_670,v200,z10,Tool_Cuy\WObj:=Workobject_1;
        MoveL Target_640,v200,z10,Tool_Cuy\WObj:=Workobject_1;
        MoveJ Target_680,v200,z10,Tool_Cuy\WObj:=Workobject_1;
        MoveJ Target_1020_3,v200,z10,Tool_Cuy\WObj:=Workobject_1;
    ENDPROC
    PROC Path_Y()
        MoveJ Target_690,v200,z10,Tool_Cuy\WObj:=Workobject_1;
        MoveL Target_700,v200,z10,Tool_Cuy\WObj:=Workobject_1;
        MoveL Target_710,v200,z10,Tool_Cuy\WObj:=Workobject_1;
        MoveL Target_720,v200,z10,Tool_Cuy\WObj:=Workobject_1;
        MoveL Target_730,v200,z10,Tool_Cuy\WObj:=Workobject_1;
        MoveL Target_740,v200,z10,Tool_Cuy\WObj:=Workobject_1;
        MoveL Target_750,v200,z10,Tool_Cuy\WObj:=Workobject_1;
        MoveL Target_760,v200,z10,Tool_Cuy\WObj:=Workobject_1;
        MoveL Target_770,v200,z10,Tool_Cuy\WObj:=Workobject_1;
        MoveL Target_690,v200,z10,Tool_Cuy\WObj:=Workobject_1;
        MoveJ Target_780,v200,z10,Tool_Cuy\WObj:=Workobject_1;
    ENDPROC
    PROC Path_E()
        MoveJ Target_790,v200,z10,Tool_Cuy\WObj:=Workobject_1;
        MoveL Target_800,v200,z10,Tool_Cuy\WObj:=Workobject_1;
        MoveL Target_810,v200,z10,Tool_Cuy\WObj:=Workobject_1;
        MoveL Target_820,v200,z10,Tool_Cuy\WObj:=Workobject_1;
        MoveL Target_830,v200,z10,Tool_Cuy\WObj:=Workobject_1;
        MoveL Target_840,v200,z10,Tool_Cuy\WObj:=Workobject_1;
        MoveL Target_850,v200,z10,Tool_Cuy\WObj:=Workobject_1;
        MoveL Target_860,v200,z10,Tool_Cuy\WObj:=Workobject_1;
        MoveL Target_870,v200,z10,Tool_Cuy\WObj:=Workobject_1;
        MoveL Target_880,v200,z10,Tool_Cuy\WObj:=Workobject_1;
        MoveL Target_890,v200,z10,Tool_Cuy\WObj:=Workobject_1;
        MoveL Target_900,v200,z10,Tool_Cuy\WObj:=Workobject_1;
        MoveL Target_790,v200,z10,Tool_Cuy\WObj:=Workobject_1;
        MoveJ Target_910,v200,z10,Tool_Cuy\WObj:=Workobject_1;
    ENDPROC
    PROC Path_I()
        MoveJ Target_920,v200,z10,Tool_Cuy\WObj:=Workobject_1;
        MoveL Target_930,v200,z10,Tool_Cuy\WObj:=Workobject_1;
        MoveL Target_940,v200,z10,Tool_Cuy\WObj:=Workobject_1;
        MoveL Target_950,v200,z10,Tool_Cuy\WObj:=Workobject_1;
        MoveL Target_920,v200,z10,Tool_Cuy\WObj:=Workobject_1;
        MoveJ Target_960,v200,z10,Tool_Cuy\WObj:=Workobject_1;
    ENDPROC
    PROC Path_S_2()
        MoveJ Target_460_2,v200,z10,Tool_Cuy\WObj:=Workobject_1;
        MoveC Target_470_2,Target_480_2,v200,z10,Tool_Cuy\WObj:=Workobject_1;
        MoveC Target_490_2,Target_500_2,v200,z10,Tool_Cuy\WObj:=Workobject_1;
        MoveL Target_510_2,v200,z10,Tool_Cuy\WObj:=Workobject_1;
        MoveC Target_520_2,Target_530_2,v200,z10,Tool_Cuy\WObj:=Workobject_1;
        MoveL Target_540_2,v200,z10,Tool_Cuy\WObj:=Workobject_1;
        MoveC Target_550_2,Target_560_2,v200,z10,Tool_Cuy\WObj:=Workobject_1;
        MoveC Target_570_2,Target_580_2,v200,z10,Tool_Cuy\WObj:=Workobject_1;
        MoveL Target_590_2,v200,z10,Tool_Cuy\WObj:=Workobject_1;
        MoveL Target_600_2,v200,z10,Tool_Cuy\WObj:=Workobject_1;
        MoveC Target_610_2,Target_620_2,v200,z10,Tool_Cuy\WObj:=Workobject_1;
        MoveL Target_460_2,v200,z10,Tool_Cuy\WObj:=Workobject_1;
        MoveJ Target_630_2,v200,z10,Tool_Cuy\WObj:=Workobject_1;
    ENDPROC
    PROC Path_O()
        MoveJ Target_970,v200,z10,Tool_Cuy\WObj:=Workobject_1;
        MoveC Target_980,Target_990,v200,z10,Tool_Cuy\WObj:=Workobject_1;
        MoveC Target_1000,Target_970,v200,z10,Tool_Cuy\WObj:=Workobject_1;
        MoveJ Target_1010,v200,z10,Tool_Cuy\WObj:=Workobject_1;
        MoveJ Target_1020,v200,z10,Tool_Cuy\WObj:=Workobject_1;
        MoveC Target_1030,Target_1040,v200,z10,Tool_Cuy\WObj:=Workobject_1;
        MoveC Target_1050,Target_1020,v200,z10,Tool_Cuy\WObj:=Workobject_1;
        MoveJ Target_1060,v200,z10,Tool_Cuy\WObj:=Workobject_1;
    ENDPROC
    PROC Path_N_2()
        MoveL Target_350_2,v1000,z100,Tool_Cuy\WObj:=Workobject_1;
        MoveL Target_360_2,v1000,z100,Tool_Cuy\WObj:=Workobject_1;
        MoveL Target_370_2,v1000,z100,Tool_Cuy\WObj:=Workobject_1;
        MoveL Target_380_2,v1000,z100,Tool_Cuy\WObj:=Workobject_1;
        MoveL Target_390_2,v1000,z100,Tool_Cuy\WObj:=Workobject_1;
        MoveL Target_400_2,v1000,z100,Tool_Cuy\WObj:=Workobject_1;
        MoveL Target_410_2,v1000,z100,Tool_Cuy\WObj:=Workobject_1;
        MoveL Target_420_2,v1000,z100,Tool_Cuy\WObj:=Workobject_1;
        MoveL Target_430_2,v1000,z100,Tool_Cuy\WObj:=Workobject_1;
        MoveL Target_440_2,v1000,z100,Tool_Cuy\WObj:=Workobject_1;
        MoveL Target_450_2,v1000,z100,Tool_Cuy\WObj:=Workobject_1;
    ENDPROC
    PROC Path_O_2()
        MoveJ Target_970_2,v200,z10,Tool_Cuy\WObj:=Workobject_1;
        MoveC Target_980_2,Target_990_2,v200,z10,Tool_Cuy\WObj:=Workobject_1;
        MoveC Target_1000_2,Target_970_2,v200,z10,Tool_Cuy\WObj:=Workobject_1;
        MoveJ Target_1010_2,v200,z10,Tool_Cuy\WObj:=Workobject_1;
        MoveJ Target_1020_2,v200,z10,Tool_Cuy\WObj:=Workobject_1;
        MoveC Target_1030_2,Target_1040_2,v200,z10,Tool_Cuy\WObj:=Workobject_1;
        MoveC Target_1050_2,Target_1020_2,v200,z10,Tool_Cuy\WObj:=Workobject_1;
        MoveJ Target_1060_2,v200,z10,Tool_Cuy\WObj:=Workobject_1;
    ENDPROC
    PROC Path_Doth_2()
        MoveJ Target_640_2,v200,z10,Tool_Cuy\WObj:=Workobject_1;
        MoveL Target_650_2,v200,z10,Tool_Cuy\WObj:=Workobject_1;
        MoveL Target_660_2,v200,z10,Tool_Cuy\WObj:=Workobject_1;
        MoveL Target_670_2,v200,z10,Tool_Cuy\WObj:=Workobject_1;
        MoveL Target_640_2,v200,z10,Tool_Cuy\WObj:=Workobject_1;
        MoveJ Target_680_2,v200,z10,Tool_Cuy\WObj:=Workobject_1;
        MoveJ Target_1020_3,v200,z10,Tool_Cuy\WObj:=Workobject_1;
    ENDPROC
    PROC Path_D()
        MoveJ Target_1070,v200,z10,Tool_Cuy\WObj:=Workobject_1;
        MoveL Target_1080,v200,z10,Tool_Cuy\WObj:=Workobject_1;
        MoveL Target_1090,v200,z10,Tool_Cuy\WObj:=Workobject_1;
        MoveC Target_1100,Target_1110,v200,z10,Tool_Cuy\WObj:=Workobject_1;
        MoveL Target_1070,v200,z10,Tool_Cuy\WObj:=Workobject_1;
        MoveJ Target_1120,v200,z10,Tool_Cuy\WObj:=Workobject_1;
        MoveJ Target_1130,v200,z10,Tool_Cuy\WObj:=Workobject_1;
        MoveL Target_1140,v200,z10,Tool_Cuy\WObj:=Workobject_1;
        MoveL Target_1150,v200,z10,Tool_Cuy\WObj:=Workobject_1;
        MoveC Target_1160,Target_1170,v200,z10,Tool_Cuy\WObj:=Workobject_1;
        MoveL Target_1130,v200,z10,Tool_Cuy\WObj:=Workobject_1;
        MoveJ Target_1180,v200,z10,Tool_Cuy\WObj:=Workobject_1;
    ENDPROC
    PROC Path_A_2()
        MoveJ Target_220_2,v200,z10,Tool_Cuy\WObj:=Workobject_1;
        MoveL Target_230_2,v200,z10,Tool_Cuy\WObj:=Workobject_1;
        MoveL Target_240_2,v200,z10,Tool_Cuy\WObj:=Workobject_1;
        MoveL Target_250_2,v200,z10,Tool_Cuy\WObj:=Workobject_1;
        MoveL Target_260_2,v200,z10,Tool_Cuy\WObj:=Workobject_1;
        MoveL Target_270_2,v200,z10,Tool_Cuy\WObj:=Workobject_1;
        MoveL Target_280_2,v200,z10,Tool_Cuy\WObj:=Workobject_1;
        MoveL Target_290_2,v200,z10,Tool_Cuy\WObj:=Workobject_1;
        MoveL Target_220_2,v200,z10,Tool_Cuy\WObj:=Workobject_1;
        MoveJ Target_300_2,v200,z10,Tool_Cuy\WObj:=Workobject_1;
        MoveJ Target_310_2,v200,z10,Tool_Cuy\WObj:=Workobject_1;
        MoveL Target_320_2,v200,z10,Tool_Cuy\WObj:=Workobject_1;
        MoveL Target_330_2,v200,z10,Tool_Cuy\WObj:=Workobject_1;
        MoveL Target_310_2,v200,z10,Tool_Cuy\WObj:=Workobject_1;
        MoveJ Target_340_2,v200,z10,Tool_Cuy\WObj:=Workobject_1;
    ENDPROC
    PROC Path_N_3()
        MoveJ Target_350_3,v200,z10,Tool_Cuy\WObj:=Workobject_1;
        MoveL Target_360_3,v200,z10,Tool_Cuy\WObj:=Workobject_1;
        MoveL Target_370_3,v200,z10,Tool_Cuy\WObj:=Workobject_1;
        MoveL Target_380_3,v200,z10,Tool_Cuy\WObj:=Workobject_1;
        MoveL Target_390_3,v200,z10,Tool_Cuy\WObj:=Workobject_1;
        MoveL Target_400_3,v200,z10,Tool_Cuy\WObj:=Workobject_1;
        MoveL Target_410_3,v200,z10,Tool_Cuy\WObj:=Workobject_1;
        MoveL Target_420_3,v200,z10,Tool_Cuy\WObj:=Workobject_1;
        MoveL Target_430_3,v200,z10,Tool_Cuy\WObj:=Workobject_1;
        MoveL Target_440_3,v200,z10,Tool_Cuy\WObj:=Workobject_1;
        MoveL Target_350_3,v200,z10,Tool_Cuy\WObj:=Workobject_1;
        MoveJ Target_450_3,v200,z10,Tool_Cuy\WObj:=Workobject_1;
    ENDPROC
    PROC Path_I_2()
        MoveJ Target_920_2,v200,z10,Tool_Cuy\WObj:=Workobject_1;
        MoveL Target_930_2,v200,z10,Tool_Cuy\WObj:=Workobject_1;
        MoveL Target_940_2,v200,z10,Tool_Cuy\WObj:=Workobject_1;
        MoveL Target_950_2,v200,z10,Tool_Cuy\WObj:=Workobject_1;
        MoveL Target_920_2,v200,z10,Tool_Cuy\WObj:=Workobject_1;
        MoveJ Target_960_2,v200,z10,Tool_Cuy\WObj:=Workobject_1;
    ENDPROC
    PROC Path_E_2()
        MoveJ Target_790_2,v200,z10,Tool_Cuy\WObj:=Workobject_1;
        MoveL Target_800_2,v200,z10,Tool_Cuy\WObj:=Workobject_1;
        MoveL Target_810_2,v200,z10,Tool_Cuy\WObj:=Workobject_1;
        MoveL Target_820_2,v200,z10,Tool_Cuy\WObj:=Workobject_1;
        MoveL Target_830_2,v200,z10,Tool_Cuy\WObj:=Workobject_1;
        MoveL Target_840_2,v200,z10,Tool_Cuy\WObj:=Workobject_1;
        MoveL Target_850_2,v200,z10,Tool_Cuy\WObj:=Workobject_1;
        MoveL Target_860_2,v200,z10,Tool_Cuy\WObj:=Workobject_1;
        MoveL Target_870_2,v200,z10,Tool_Cuy\WObj:=Workobject_1;
        MoveL Target_880_2,v200,z10,Tool_Cuy\WObj:=Workobject_1;
        MoveL Target_890_2,v200,z10,Tool_Cuy\WObj:=Workobject_1;
        MoveL Target_900_2,v200,z10,Tool_Cuy\WObj:=Workobject_1;
        MoveL Target_790_2,v200,z10,Tool_Cuy\WObj:=Workobject_1;
        MoveJ Target_910_2,v200,z10,Tool_Cuy\WObj:=Workobject_1;
    ENDPROC
    PROC Path_L()
        MoveJ Target_1190,v200,z10,Tool_Cuy\WObj:=Workobject_1;
        MoveL Target_1200,v200,z10,Tool_Cuy\WObj:=Workobject_1;
        MoveL Target_1210,v200,z10,Tool_Cuy\WObj:=Workobject_1;
        MoveL Target_1220,v200,z10,Tool_Cuy\WObj:=Workobject_1;
        MoveL Target_1230,v200,z10,Tool_Cuy\WObj:=Workobject_1;
        MoveL Target_1240,v200,z10,Tool_Cuy\WObj:=Workobject_1;
        MoveL Target_1190,v200,z10,Tool_Cuy\WObj:=Workobject_1;
        MoveJ Target_1250,v200,z10,Tool_Cuy\WObj:=Workobject_1;
    ENDPROC
    PROC Path_R()
        MoveJ Target_1260,v200,z10,Tool_Cuy\WObj:=Workobject_1;
        MoveL Target_1270,v200,z10,Tool_Cuy\WObj:=Workobject_1;
        MoveL Target_1280,v200,z10,Tool_Cuy\WObj:=Workobject_1;
        MoveL Target_1290,v200,z10,Tool_Cuy\WObj:=Workobject_1;
        MoveL Target_1300,v200,z10,Tool_Cuy\WObj:=Workobject_1;
        MoveC Target_1310,Target_1320,v200,z10,Tool_Cuy\WObj:=Workobject_1;
        MoveL Target_1330,v200,z10,Tool_Cuy\WObj:=Workobject_1;
        MoveL Target_1340,v200,z10,Tool_Cuy\WObj:=Workobject_1;
        MoveL Target_1350,v200,z10,Tool_Cuy\WObj:=Workobject_1;
        MoveC Target_1360,Target_1370,v200,z10,Tool_Cuy\WObj:=Workobject_1;
        MoveL Target_1380,v200,z10,Tool_Cuy\WObj:=Workobject_1;
        MoveC Target_1390,Target_1400,v200,z10,Tool_Cuy\WObj:=Workobject_1;
        MoveL Target_1260,v200,z10,Tool_Cuy\WObj:=Workobject_1;
        MoveJ Target_1410,v200,z10,Tool_Cuy\WObj:=Workobject_1;
        MoveJ Target_1420,v200,z10,Tool_Cuy\WObj:=Workobject_1;
        MoveL Target_1430,v200,z10,Tool_Cuy\WObj:=Workobject_1;
        MoveL Target_1440,v200,z10,Tool_Cuy\WObj:=Workobject_1;
        MoveC Target_1450,Target_1460,v200,z10,Tool_Cuy\WObj:=Workobject_1;
        MoveL Target_1420,v200,z10,Tool_Cuy\WObj:=Workobject_1;
        MoveJ Target_1470,v200,z10,Tool_Cuy\WObj:=Workobject_1;
    ENDPROC
    PROC Path_Doth_3()
        MoveJ Target_640_3,v200,z10,Tool_Cuy\WObj:=Workobject_1;
        MoveL Target_650_3,v200,z10,Tool_Cuy\WObj:=Workobject_1;
        MoveL Target_660_3,v200,z10,Tool_Cuy\WObj:=Workobject_1;
        MoveL Target_670_3,v200,z10,Tool_Cuy\WObj:=Workobject_1;
        MoveL Target_640_3,v200,z10,Tool_Cuy\WObj:=Workobject_1;
        MoveJ Target_680_3,v200,z10,Tool_Cuy\WObj:=Workobject_1;
        MoveJ Target_1020_3,v200,z10,Tool_Cuy\WObj:=Workobject_1;
    ENDPROC
    PROC Path_Cuy_Externo()
        MoveJ Target_1480,v200,z10,Tool_Cuy\WObj:=Workobject_1;
        MoveC Target_1490,Target_1500,v200,z10,Tool_Cuy\WObj:=Workobject_1;
        MoveC Target_1510,Target_1520,v200,z10,Tool_Cuy\WObj:=Workobject_1;
        MoveL Target_1530,v200,z10,Tool_Cuy\WObj:=Workobject_1;
        MoveC Target_1540,Target_1550,v200,z10,Tool_Cuy\WObj:=Workobject_1;
        MoveC Target_1560,Target_1580,v200,z10,Tool_Cuy\WObj:=Workobject_1;
        MoveC Target_1590,Target_1600,v200,z10,Tool_Cuy\WObj:=Workobject_1;
        MoveL Target_1610,v200,z10,Tool_Cuy\WObj:=Workobject_1;
        MoveC Target_1620,Target_1640,v200,z10,Tool_Cuy\WObj:=Workobject_1;
        MoveL Target_1650,v200,z10,Tool_Cuy\WObj:=Workobject_1;
        MoveC Target_1660,Target_1670,v200,z10,Tool_Cuy\WObj:=Workobject_1;
        MoveL Target_1680,v200,z10,Tool_Cuy\WObj:=Workobject_1;
        MoveC Target_1690,Target_1700,v200,z10,Tool_Cuy\WObj:=Workobject_1;
        MoveL Target_1710,v200,z10,Tool_Cuy\WObj:=Workobject_1;
        MoveL Target_1720,v200,z10,Tool_Cuy\WObj:=Workobject_1;
        MoveC Target_1730,Target_1740,v200,z10,Tool_Cuy\WObj:=Workobject_1;
        MoveC Target_1750,Target_1760,v200,z10,Tool_Cuy\WObj:=Workobject_1;
        MoveL Target_1770,v200,z10,Tool_Cuy\WObj:=Workobject_1;
        MoveC Target_1780,Target_1790,v200,z10,Tool_Cuy\WObj:=Workobject_1;
        MoveC Target_1800,Target_1810,v200,z10,Tool_Cuy\WObj:=Workobject_1;
        MoveL Target_1480,v200,z10,Tool_Cuy\WObj:=Workobject_1;
        MoveJ Target_1820,v200,z10,Tool_Cuy\WObj:=Workobject_1;
    ENDPROC
    PROC Path_Cuy_Interno()
        MoveJ Target_1830,v200,z10,Tool_Cuy\WObj:=Workobject_1;
        MoveC Target_1840,Target_1850,v200,z10,Tool_Cuy\WObj:=Workobject_1;
        MoveL Target_1860,v200,z10,Tool_Cuy\WObj:=Workobject_1;
        MoveC Target_1870,Target_1880,v200,z10,Tool_Cuy\WObj:=Workobject_1;
        MoveL Target_1900,v200,z10,Tool_Cuy\WObj:=Workobject_1;
        MoveC Target_1910,Target_1920,v200,z10,Tool_Cuy\WObj:=Workobject_1;
        MoveL Target_1930,v200,z10,Tool_Cuy\WObj:=Workobject_1;
        MoveC Target_1940,Target_1950,v200,z10,Tool_Cuy\WObj:=Workobject_1;
        MoveC Target_1960,Target_1970,v200,z10,Tool_Cuy\WObj:=Workobject_1;
        MoveL Target_1980,v200,z10,Tool_Cuy\WObj:=Workobject_1;
        MoveC Target_2000,Target_2010,v200,z10,Tool_Cuy\WObj:=Workobject_1;
        MoveL Target_2020,v200,z10,Tool_Cuy\WObj:=Workobject_1;
        MoveL Target_2040,v200,z10,Tool_Cuy\WObj:=Workobject_1;
        MoveC Target_2050,Target_2060,v200,z10,Tool_Cuy\WObj:=Workobject_1;
        MoveL Target_2080,v200,z10,Tool_Cuy\WObj:=Workobject_1;
        MoveC Target_2090,Target_2100,v200,z10,Tool_Cuy\WObj:=Workobject_1;
        MoveL Target_2110,v200,z10,Tool_Cuy\WObj:=Workobject_1;
        MoveL Target_2120,v200,z10,Tool_Cuy\WObj:=Workobject_1;
        MoveC Target_2130,Target_2140,v200,z10,Tool_Cuy\WObj:=Workobject_1;
        MoveC Target_2150,Target_2160,v200,z10,Tool_Cuy\WObj:=Workobject_1;
        MoveC Target_2170,Target_2180,v200,z10,Tool_Cuy\WObj:=Workobject_1;
        MoveC Target_2190,Target_2200,v200,z10,Tool_Cuy\WObj:=Workobject_1;
        MoveC Target_2220,Target_1830,v200,z10,Tool_Cuy\WObj:=Workobject_1;
        MoveJ Target_2210,v200,z10,Tool_Cuy\WObj:=Workobject_1;
    ENDPROC
    PROC Path_Oreja()
        MoveJ Target_2230,v200,z10,Tool_Cuy\WObj:=Workobject_1;
        MoveC Target_2240,Target_2250,v200,z10,Tool_Cuy\WObj:=Workobject_1;
        MoveC Target_2260,Target_2270,v200,z10,Tool_Cuy\WObj:=Workobject_1;
        MoveC Target_2280,Target_2290,v200,z10,Tool_Cuy\WObj:=Workobject_1;
        MoveJ Target_2300,v200,z10,Tool_Cuy\WObj:=Workobject_1;
    ENDPROC
    PROC Path_Ojo()
        MoveJ Target_2310,v200,z10,Tool_Cuy\WObj:=Workobject_1;
        MoveC Target_2320,Target_2330,v200,z10,Tool_Cuy\WObj:=Workobject_1;
        MoveC Target_2340,Target_2310,v200,z10,Tool_Cuy\WObj:=Workobject_1;
        MoveJ Target_2350,v200,z10,Tool_Cuy\WObj:=Workobject_1;
    ENDPROC
    PROC FarmearAura()
        Path_Home;
        ! Posición inicial erguida
        MoveAbsJ Aura_Vertical,v800,fine,Tool_Cuy;

        ! Empieza a abrirse mientras gira
        MoveAbsJ Aura_Abre_Der,v400,z10,Tool_Cuy;
        MoveAbsJ Aura_Giro_Der,v400,z10,Tool_Cuy;

        ! Giro hacia el lado contrario
        MoveAbsJ Aura_Abre_Izq,v800,z10,Tool_Cuy;
        MoveAbsJ Aura_Giro_Izq,v800,z10,Tool_Cuy;

        ! Segunda vuelta más rápida
        MoveAbsJ Aura_Giro_Der,v400,z10,Tool_Cuy;
        MoveAbsJ Aura_Giro_Izq,v400,z10,Tool_Cuy;

        ! Cierre elegante
        MoveAbsJ Aura_Abre_Der,v800,z20,Tool_Cuy;
        MoveAbsJ Aura_Vertical,v800,fine,Tool_Cuy;

        ! Saludo rápido con muñeca
        MoveAbsJ Aura_Saludo_1,v1000,z10,Tool_Cuy;
        MoveAbsJ Aura_Saludo_2,v1000,z10,Tool_Cuy;
        MoveAbsJ Aura_Saludo_3,v1000,z10,Tool_Cuy;
        MoveAbsJ Aura_Saludo_4,v1000,z10,Tool_Cuy;
        MoveAbsJ Aura_Saludo_5,v1000,z10,Tool_Cuy;
        MoveAbsJ Aura_Saludo_6,v1000,z10,Tool_Cuy;
        MoveAbsJ Aura_Saludo_Fin,v1000,fine,Tool_Cuy;

        Path_Home;
    ENDPROC
    PROC Mantenimiento()
        Path_Home;
        MoveAbsJ Mant_Aprox,v400,fine,Tool_Cuy;

    ENDPROC

ENDMODULE
